// TwinCAT 3 PLC project PLC_Dyno
// ProgramVersion: 3.1.4026.25
// CompilerDefines: VISU_USEPROPERTYINFO
// libraries:
//   CmpBitmapPool, * (System)
//   Tc2_EtherCAT, * (Beckhoff Automation GmbH)
//   Tc2_MC2, * (Beckhoff Automation GmbH)
//   Tc2_MC2_Drive, * (Beckhoff Automation GmbH)
//   Tc2_Standard, * (Beckhoff Automation GmbH)
//   Tc2_System, * (Beckhoff Automation GmbH)
//   VisuDialogs, * (System)
//   VisuSymbols, 4.5.0.0 (System)
// project tree:
//   DUTs/ E_ControlMode.TcDUT, E_MotorState.TcDUT, E_SafetyState.TcTLEO, ST_AnalogInData.TcDUT, ST_EncoderData.TcDUT, ST_IOData.TcDUT, ST_MenteeMotorCmd.TcDUT, ST_MenteeMotorStatus.TcDUT, ST_MenteeMotorV32OsCmd.TcDUT, ST_MenteeMotorV32OsSample.TcDUT, ST_MenteeMotorV32OsStatus.TcDUT, ST_MenteeTrajCmd.TcDUT, ST_LoadProfileCmd.TcDUT, ST_CsvProfile.TcDUT, ST_Slot2Cfg.TcDUT, ST_MotorCommand.TcDUT, ST_RecChunk.TcDUT, U_WordReal.TcDUT, ST_MotorStatus.TcDUT, ST_Safety_Speps.TcDUT, ST_SyncSnapshot.TcDUT, ST_TwinSAFE_IN.TcDUT, ST_TwinSAFE_OUT.TcDUT, ST_UartBridgeCmd.TcDUT, ST_UartBridgeStatus.TcDUT
//   / GlobalTextList.TcGTLO, ImagePool.TcIPO (not stored), PlcTask.TcTTO, Visualization Manager.TcVMO (not stored), VISU_TASK.TcTTO
//   GVLs/ GVL_AnalogIn.TcGVL, GVL_Commands.TcGVL, GVL_MenteeFoe.TcGVL, GVL_Encoder.TcGVL, GVL_IO.TcGVL, GVL_MenteeMotor.TcGVL, GVL_MenteeMotorV32_OS.TcGVL, GVL_Profiles.TcGVL, GVL_CsvProfile.TcGVL, GVL_Slot2.TcGVL, GVL_Recording.TcGVL, GVL_Safety.TcGVL, GVL_Status.TcGVL, GVL_Sync.TcGVL, GVL_UartBridge.TcGVL
//   POUs/ CheckBounds.TcPOU, FB_AnalogInHandler.TcPOU, FB_EncoderHandler.TcPOU, FB_IOHandler.TcPOU, FB_MenteeMotorHandler.TcPOU, FB_MotorControl.TcPOU, FB_ExtSetpointProbe.TcPOU, FB_LoadMotorProfile.TcPOU, FB_CsvPlayer.TcPOU, FB_MenteeSdoCmd.TcPOU, FB_MenteeFoeFlash.TcPOU, FB_Slot2PipeHandler.TcPOU, FB_TorqueControl.TcPOU, FB_HighRateRecorder.TcPOU, FB_TrajectoryGen.TcPOU, FB_UartBridgeHandler.TcPOU, MAIN.TcPOU, PRG_Motion.TcPOU
//   VISUs/ Visualization.TcVIS
// real-time tasks:
//   TASK PlcTask: cycle T#1ms, priority 2, ADS port 350
//   TASK VISU_TASK: cycle T#200000us, priority 30, ADS port 351
// motion (NC):
//   TASK NC-Task 1 SAF: cycle T#1ms, priority 4, ADS port 501
//   TASK NC-Task 1 SVB: cycle T#10ms, priority 8, ADS port 511
//   AXIS Axis 1 (id 3)
//     General: UnitName=°
//     Dynamic: Acceleration=15000, Deceleration=15000, Jerk=178490.844
//     Velo: RefSearch=396.64632, RefSync=396.64632, SlowManual=1983.2316, FastManual=11899.3896, Fast=39664.632, Maximum=39664.632
//     OtherSettings: AllowMotionCmdToSlave=true
//     encoder EncType=8
//       EncPara: ScaleFactorNumerator=360, ScaleFactorDenominator=1048576, MaxCount=#xffffffff, EncPositionSource=1
//     drive DrvType=9
//       DrvPara: MaxCount=#xffffffff, DriveControlDWord=#x00030100
//         Analog: VeloReferenz=43631.0952, VeloScale=1.02400649589962, TorqueSetpointScale=10, ScaleFactorActTorque=0.1
//         TimeComp: TaskDelayCycles=1
//     controller CtrType=1
//       CtrPara: PriorControlFactor=1
//         Observer: BandWidth=20
//   AXIS Axis 2 (id 4)
//     General: UnitName=°
//     Dynamic: Acceleration=13437.441, Deceleration=13437.441, Jerk=40312.323
//     Velo: RefSearch=89.58294, RefSync=89.58294, SlowManual=447.9147, FastManual=2687.4882, Fast=8958.294, Maximum=8958.294
//     OtherSettings: AllowMotionCmdToSlave=true
//     encoder EncType=8
//       EncPara: ScaleFactorNumerator=360, ScaleFactorDenominator=1048576, MaxCount=#xffffffff
//     drive DrvType=9
//       DrvPara: MaxCount=#xffffffff, DriveControlDWord=#x00030100
//         Analog: VeloReferenz=9854.1234, VeloScale=1.02400649589962, TorqueSetpointScale=10, ScaleFactorActTorque=0.1
//         TimeComp: TaskDelayCycles=1
//     controller CtrType=1
//       CtrPara: PriorControlFactor=1
//         Observer: BandWidth=20
// I/O:
//   DEVICE Device 2 (EtherCAT), AmsNetId 192.168.1.50.3.1
//     Machine Side - A10 (EK1200)_1 [EK1200-5000 EtherCAT Power supply (2A E-Bus)]
//       A11 - DO (EL2022)_1 [EL2022 2Ch. Dig. Output 24V, 2A]
//       Term 3 (EL2502) [EL2502 2Ch. PWM output, 24V]
//       A12 - SI2 (EL1918)_1 [EL1918, 8Ch. Safety Input 24V, TwinSAFE]
//         modules: Module 1 (FSOE), Module 2 (FSLOGIC)
//       A13 - SO3 (EL2904)_1 [EL2904, 4 Ch. Safety Output 24V, 0.5A, TwinSAFE]
//         modules: Module 1 (FSOES), Module 2 (DO)
//       A14 - D-I/O (EL1859)_1 [EL1859 8Ch. Dig. Input 24V, 3ms, 8Ch. Dig. Output 24V, 0.5A]
//       A15 - AI (EL3002)_1 [EL3002 2Ch. Ana. Input +/-10V]
//       A19 - Enc (EL5112)_1 [EL5112 2Ch. Inc. Encoder 5V (2xAB or 1xABC RS422,TTL)]
//       A16 - AI  (EL3702)_1 [EL3702 2Ch. Ana. Input +/-10V, DIFF, Oversample]
//       A18 - Enc  (EL5112)_1 [EL5112 2Ch. Inc. Encoder 5V (2xAB or 1xABC RS422,TTL)]
//       A17 - AI  (EL3702)_1 [EL3702 2Ch. Ana. Input +/-10V, DIFF, Oversample]
//       Term 12 (EL5042) [EL5042 2Ch. BiSS-C Encoder]
//       Term 14 (EK1110)_1 [EK1110 EtherCAT extension]
//     Drive 1 (AX5112-0000-0216) [AX5112-0000-0216 EtherCAT Drive (SoE, 1 Ch.)]
//       STO_Drive1 (AX5805) [AX5805 (Safety Drive Option)]
//         modules: Module 1 (Safety Process Data, 1 axis), Module 2 (Standard Process Data, 1 axis)
//     Drive 2 (AX5125-0000-0216) [AX5125-0000-0216 EtherCAT Drive (SoE, 1 Ch.)]
//       STO_Drive2 (AX5805) [AX5805 (Safety Drive Option)]
//         modules: Module 1 (Safety Process Data, 1 axis), Module 2 (Standard Process Data, 1 axis)
//     Rack 19 (EK1100 - A0)_1 [EK1100 EtherCAT Coupler (2A E-Bus)]
//       A1 - SI1 (EL1918)_1 [EL1918, 8Ch. Safety Input 24V, TwinSAFE]
//         modules: Module 2 (FSLOGIC)
//       A2 -SO1 (EL2904)_1 [EL2904, 4 Ch. Safety Output 24V, 0.5A, TwinSAFE]
//         modules: Module 1 (FSOES), Module 2 (DO)
//       A3 - SO2 (EL2904)_1 [EL2904, 4 Ch. Safety Output 24V, 0.5A, TwinSAFE]
//         modules: Module 1 (FSOES), Module 2 (DO)
//       A4 - D-I/O (EL1859)_1 [EL1859 8Ch. Dig. Input 24V, 3ms, 8Ch. Dig. Output 24V, 0.5A]
//       A5 (EL9505)_1 [EL9505 Power supply terminal 5V]
//       A6  (EL9505)_1 [EL9505 Power supply terminal 5V]
//       Term 23 (EL9011) [EL9011 End Terminal]
//     Box 1 (Motor Slave) [Motor Slave]
// variable links:
//   Device 2 (EtherCAT) <-> Device 2 (EtherCAT)/Rack 19 (EK1100 - A0)_1/A1 - SI1 (EL1918)_1
//     Drive 1 (AX5112-0000-0216)/STO_Drive1 (AX5805)/Module 1 (Safety Process Data, 1 axis)/Inputs (Statusword)/FSOE <-> ConnectionOutputs/Message_71 RxPDO
//     Drive 2 (AX5125-0000-0216)/STO_Drive2 (AX5805)/Module 1 (Safety Process Data, 1 axis)/Inputs (Statusword)/FSOE <-> ConnectionOutputs/Message_72 RxPDO
//     Drive 1 (AX5112-0000-0216)/STO_Drive1 (AX5805)/Module 1 (Safety Process Data, 1 axis)/Outputs (Controlword)/FSOE <-> ConnectionInputs/Message_71 TxPDO
//     Drive 2 (AX5125-0000-0216)/STO_Drive2 (AX5805)/Module 1 (Safety Process Data, 1 axis)/Outputs (Controlword)/FSOE <-> ConnectionInputs/Message_72 TxPDO
//     Machine Side - A10 (EK1200)_1/A12 - SI2 (EL1918)_1/Module 1 (FSOE)/FSoE Inputs/FSOE <-> ConnectionOutputs/Message_62 RxPDO
//     Machine Side - A10 (EK1200)_1/A12 - SI2 (EL1918)_1/Module 1 (FSOE)/FSoE Outputs/FSOE <-> ConnectionInputs/Message_62 TxPDO
//     Machine Side - A10 (EK1200)_1/A13 - SO3 (EL2904)_1/Module 1 (FSOES)/RxPDO/FSOE <-> ConnectionInputs/Message_51 TxPDO
//     Machine Side - A10 (EK1200)_1/A13 - SO3 (EL2904)_1/Module 1 (FSOES)/TxPDO/FSOE <-> ConnectionOutputs/Message_51 RxPDO
//   Device 2 (EtherCAT) <-> Device 2 (EtherCAT)/Rack 19 (EK1100 - A0)_1/A2 -SO1 (EL2904)_1
//     Rack 19 (EK1100 - A0)_1/A1 - SI1 (EL1918)_1/ConnectionInputs/Message_7 TxPDO <-> Module 1 (FSOES)/RxPDO/FSOE
//     Rack 19 (EK1100 - A0)_1/A1 - SI1 (EL1918)_1/ConnectionOutputs/Message_7 RxPDO <-> Module 1 (FSOES)/TxPDO/FSOE
//   Device 2 (EtherCAT) <-> Device 2 (EtherCAT)/Rack 19 (EK1100 - A0)_1/A3 - SO2 (EL2904)_1
//     Rack 19 (EK1100 - A0)_1/A1 - SI1 (EL1918)_1/ConnectionInputs/Message_8 TxPDO <-> Module 1 (FSOES)/RxPDO/FSOE
//     Rack 19 (EK1100 - A0)_1/A1 - SI1 (EL1918)_1/ConnectionOutputs/Message_8 RxPDO <-> Module 1 (FSOES)/TxPDO/FSOE
//   NC-Task 1 SAF/Axes/Axis 1 <-> Device 2 (EtherCAT)/Drive 1 (AX5112-0000-0216)
//     Drive/Inputs/In/nDataIn1 <-> AT/Following distance
//     Drive/Inputs/In/nDataIn3[0] <-> AT/Torque/force feedback value
//     Drive/Inputs/In/nDcOutputTime <-> InfoData/DcOutputShift
//     Drive/Inputs/In/nState1 <-> AT/Drive status word @bit 8
//     Drive/Inputs/In/nState2 <-> AT/Drive status word
//     Drive/Inputs/In/nState4 @bit 1 <-> WcState/InputToggle
//     Drive/Inputs/In/nState4 <-> WcState/WcState
//     Drive/Outputs/Out/nCtrl1 <-> MDT/Master control word @bit 8
//     Drive/Outputs/Out/nDataOut1 <-> MDT/Position command value
//     Drive/Outputs/Out/nDataOut4[0] <-> MDT/Torque/force command value
//     Drive/Outputs/Out/nDataOut5 <-> MDT/High velocity limit value
//     Drive/Outputs/Out/nDataOut6 <-> MDT/Low velocity limit value
//     Enc/Inputs/In/nDataIn1 <-> AT/Position feedback 1 value
//     Enc/Inputs/In/nDataIn7 <-> AT/Velocity feedback 1 value
//     Enc/Inputs/In/nDcInputTime <-> InfoData/DcInputShift
//     Enc/Inputs/In/nState4 @bit 1 <-> WcState/InputToggle
//     Enc/Inputs/In/nState4 <-> WcState/WcState
//   NC-Task 1 SAF/Axes/Axis 2 <-> Device 2 (EtherCAT)/Drive 2 (AX5125-0000-0216)
//     Drive/Inputs/In/nDataIn1 <-> AT/Following distance
//     Drive/Inputs/In/nDcOutputTime <-> InfoData/DcOutputShift
//     Drive/Inputs/In/nState1 <-> AT/Drive status word @bit 8
//     Drive/Inputs/In/nState2 <-> AT/Drive status word
//     Drive/Inputs/In/nState4 @bit 1 <-> WcState/InputToggle
//     Drive/Inputs/In/nState4 <-> WcState/WcState
//     Drive/Outputs/Out/nCtrl1 <-> MDT/Master control word @bit 8
//     Drive/Outputs/Out/nDataOut1 <-> MDT/Position command value
//     Drive/Outputs/Out/nDataOut4[0] <-> MDT/Torque/force command value
//     Drive/Outputs/Out/nDataOut5 <-> MDT/High velocity limit value
//     Drive/Outputs/Out/nDataOut6 <-> MDT/Low velocity limit value
//     Enc/Inputs/In/nDataIn1 <-> AT/Position feedback 1 value
//     Enc/Inputs/In/nDcInputTime <-> InfoData/DcInputShift
//     Enc/Inputs/In/nState4 @bit 1 <-> WcState/InputToggle
//     Enc/Inputs/In/nState4 <-> WcState/WcState
//   PLC_Dyno/PLC_Dyno Instance <-> Device 2 (EtherCAT)/Box 1 (Motor Slave)
//     PlcTask Inputs/GVL_MenteeMotorV32_OS.nSlaveState <-> InfoData/State
//     PlcTask Inputs/PRG_Motion.fbMenteeSdo.stAdsAddr <-> InfoData/AdsAddr
//     PlcTask Inputs/PRG_Motion.fbSlot2Pipe.i_capture_count <-> Motor Response TB/capture_count
//     PlcTask Inputs/PRG_Motion.fbSlot2Pipe.i_categorial_error <-> Motor Response TB/categorial_error
//     PlcTask Inputs/PRG_Motion.fbSlot2Pipe.i_fault <-> Motor Response TB/fault
//     PlcTask Inputs/PRG_Motion.fbSlot2Pipe.i_fsm_state <-> Motor Response TB/fsm_state
//     PlcTask Inputs/PRG_Motion.fbSlot2Pipe.i_general_error <-> Motor Response TB/general_error
//     PlcTask Inputs/PRG_Motion.fbSlot2Pipe.i_last_op <-> Motor Response TB/last_op
//     PlcTask Inputs/PRG_Motion.fbSlot2Pipe.i_main_state <-> Motor Response TB/main_state
//     PlcTask Inputs/PRG_Motion.fbSlot2Pipe.i_motion_mode <-> Motor Response TB/motion_mode
//     PlcTask Inputs/PRG_Motion.fbSlot2Pipe.i_motor_enabled <-> Motor Response TB/motor_enabled
//     PlcTask Inputs/PRG_Motion.fbSlot2Pipe.i_sample_count <-> Motor Response TB/sample_count
//     PlcTask Inputs/PRG_Motion.fbSlot2Pipe.i_samples[{0..99}] <-> Motor Response TB/sample_{0..99}  (100 links)
//     PlcTask Inputs/PRG_Motion.fbSlot2Pipe.i_var_count <-> Motor Response TB/var_count
//     PlcTask Outputs/PRG_Motion.fbSlot2Pipe.q_addr <-> Motor Command TB/addr_payload
//     PlcTask Outputs/PRG_Motion.fbSlot2Pipe.q_inject[{0..9}] <-> Motor Command TB/inject_{0..9}  (10 links)
//     PlcTask Outputs/PRG_Motion.fbSlot2Pipe.q_op <-> Motor Command TB/op
//     PlcTask Outputs/PRG_Motion.fbSlot2Pipe.q_prescaler <-> Motor Command TB/prescaler
//     PlcTask Outputs/PRG_Motion.fbSlot2Pipe.q_size <-> Motor Command TB/size
//     PlcTask Outputs/PRG_Motion.fbSlot2Pipe.q_slot <-> Motor Command TB/slot
//     PlcTask Outputs/PRG_Motion.fbSlot2Pipe.q_strobe <-> Motor Command TB/strobe
//   PLC_Dyno/PLC_Dyno Instance <-> Device 2 (EtherCAT)/Drive 1 (AX5112-0000-0216)
//     PlcTask Inputs/PRG_Motion.fbMotor1.nActTorque_Raw <-> AT/Torque/force feedback value
//     PlcTask Outputs/GVL_Commands.nMotor1_CurrentLimit_Raw <-> MDT/Bipolar torque/force limit value
//   PLC_Dyno/PLC_Dyno Instance <-> Device 2 (EtherCAT)/Drive 2 (AX5125-0000-0216)
//     PlcTask Inputs/PRG_Motion.fbMotor2.nActTorque_Raw <-> AT/Torque/force feedback value
//     PlcTask Outputs/GVL_Commands.nMotor2_CurrentLimit_Raw <-> MDT/Bipolar torque/force limit value
//   PLC_Dyno/PLC_Dyno Instance <-> Device 2 (EtherCAT)/Machine Side - A10 (EK1200)_1/A14 - D-I/O (EL1859)_1
//     PlcTask Inputs/GVL_Safety.DoorMonitorFromPLC <-> Channel 2/Input
//     PlcTask Inputs/GVL_Safety.SolonoidStatus <-> Channel 1/Input
//     PlcTask Outputs/GVL_IO.BlueLED <-> Channel 11/Output
//     PlcTask Outputs/GVL_IO.GreenLED <-> Channel 10/Output
//     PlcTask Outputs/GVL_IO.RedLED <-> Channel 9/Output
//     PlcTask Outputs/GVL_IO.b_MotorCooling <-> Channel 12/Output
//   PLC_Dyno/PLC_Dyno Instance <-> Device 2 (EtherCAT)/Machine Side - A10 (EK1200)_1/A16 - AI  (EL3702)_1
//     PlcTask Inputs/PRG_Motion.fbAnalogIn1.nCh1_S{1..5} <-> Ch1 Sample {0..4}/Ch1 Value  (5 links)
//   PLC_Dyno/PLC_Dyno Instance <-> Device 2 (EtherCAT)/Machine Side - A10 (EK1200)_1/A17 - AI  (EL3702)_1
//     PlcTask Inputs/PRG_Motion.fbAnalogIn2.nCh1_S{1..5} <-> Ch1 Sample {0..4}/Ch1 Value  (5 links)
//   PLC_Dyno/PLC_Dyno Instance <-> Device 2 (EtherCAT)/Machine Side - A10 (EK1200)_1/A18 - Enc  (EL5112)_1
//     PlcTask Inputs/PRG_Motion.fbEncoder2.nCounterValue_Raw <-> ENC Status Channel 1/Counter value
//     PlcTask Inputs/PRG_Motion.fbEncoder2.nFrequencyValue_Raw <-> ENC Frequency Channel 1/Frequency value
//     PlcTask Outputs/PRG_Motion.fbEncoder2.nControlWord_Raw <-> ENC Control Channel 1/Control
//     PlcTask Outputs/PRG_Motion.fbEncoder2.nSetCounterValue_Raw <-> ENC Control Channel 1/Set counter value
//   PLC_Dyno/PLC_Dyno Instance <-> Device 2 (EtherCAT)/Machine Side - A10 (EK1200)_1/A19 - Enc (EL5112)_1
//     PlcTask Inputs/PRG_Motion.fbEncoder1.nCounterValue_Raw <-> ENC Status Channel 1/Counter value
//     PlcTask Inputs/PRG_Motion.fbEncoder1.nFrequencyValue_Raw <-> ENC Frequency Channel 1/Frequency value
//     PlcTask Outputs/PRG_Motion.fbEncoder1.nControlWord_Raw <-> ENC Control Channel 1/Control
//     PlcTask Outputs/PRG_Motion.fbEncoder1.nSetCounterValue_Raw <-> ENC Control Channel 1/Set counter value
//   PLC_Dyno/PLC_Dyno Instance <-> Device 2 (EtherCAT)/Rack 19 (EK1100 - A0)_1/A1 - SI1 (EL1918)_1
//     PlcTask Inputs/GVL_Safety.stTwinSAFE_IN/C1_FBK <-> StandardInputs/Standard Out Var 87
//     PlcTask Inputs/GVL_Safety.stTwinSAFE_IN/C2_FBK <-> StandardInputs/Standard Out Var 88
//     PlcTask Inputs/GVL_Safety.stTwinSAFE_IN/EStop_MantiRob <-> StandardInputs/Standard Out Var 84
//     PlcTask Inputs/GVL_Safety.stTwinSAFE_IN/EStop_NC1 <-> StandardInputs/Standard Out Var 82
//     PlcTask Inputs/GVL_Safety.stTwinSAFE_IN/EStop_NC2 <-> StandardInputs/Standard Out Var 83
//     PlcTask Inputs/GVL_Safety.stTwinSAFE_IN/EStop_Ok <-> StandardInputs/Standard Out Var 77
//     PlcTask Inputs/GVL_Safety.stTwinSAFE_IN/EStop_Status <-> StandardInputs/Standard Out Var 78
//     PlcTask Inputs/GVL_Safety.stTwinSAFE_IN/HV_Healthy <-> StandardInputs/Standard Out Var 90
//     PlcTask Inputs/GVL_Safety.stTwinSAFE_IN/HV_Interlock <-> StandardInputs/Standard Out Var 92
//     PlcTask Inputs/GVL_Safety.stTwinSAFE_IN/LV_Healthy <-> StandardInputs/Standard Out Var 89
//     PlcTask Inputs/GVL_Safety.stTwinSAFE_IN/LV_Interlock <-> StandardInputs/Standard Out Var 91
//     PlcTask Inputs/GVL_Safety.stTwinSAFE_IN/ReadyForStep2 <-> StandardInputs/Standard Out Var 52
//     PlcTask Inputs/GVL_Safety.stTwinSAFE_IN/STO_1 <-> StandardInputs/Standard Out Var 85
//     PlcTask Inputs/GVL_Safety.stTwinSAFE_IN/STO_2 <-> StandardInputs/Standard Out Var 86
//     PlcTask Inputs/GVL_Safety.stTwinSAFE_IN/Safety_Armed <-> StandardInputs/Standard Out Var 53
//     PlcTask Inputs/GVL_Safety.stTwinSAFE_IN/Speps/step{1..6} <-> StandardInputs/Standard Out Var {65..70}  (6 links)
//     PlcTask Inputs/GVL_Safety.stTwinSAFE_IN/Speps/stepRnD <-> StandardInputs/Standard Out Var 95
//     PlcTask Inputs/GVL_Safety.stTwinSAFE_IN/TransitionStep <-> StandardInputs/Standard Out Var 98
//     PlcTask Outputs/GVL_Safety.stTwinSAFE_OUT/BatRelay_Manual_Off <-> StandardOutputs/Standard In Var 56
//     PlcTask Outputs/GVL_Safety.stTwinSAFE_OUT/BatRelay_Manual_On <-> StandardOutputs/Standard In Var 55
//     PlcTask Outputs/GVL_Safety.stTwinSAFE_OUT/Bypass_C1C2 <-> StandardOutputs/Standard In Var 99
//     PlcTask Outputs/GVL_Safety.stTwinSAFE_OUT/DoorMonitor <-> StandardOutputs/Standard In Var 16
//     PlcTask Outputs/GVL_Safety.stTwinSAFE_OUT/ErrACK <-> StandardOutputs/Standard In Var 1
//     PlcTask Outputs/GVL_Safety.stTwinSAFE_OUT/EstopPLC <-> StandardOutputs/Standard In Var 54
//     PlcTask Outputs/GVL_Safety.stTwinSAFE_OUT/RB_BatBMS_Manual_Off <-> StandardOutputs/Standard In Var 58
//     PlcTask Outputs/GVL_Safety.stTwinSAFE_OUT/RB_BatBMS_Manual_On <-> StandardOutputs/Standard In Var 57
//     PlcTask Outputs/GVL_Safety.stTwinSAFE_OUT/RUN <-> StandardOutputs/Standard In Var 50
//     PlcTask Outputs/GVL_Safety.stTwinSAFE_OUT/Set_RnD_Mode <-> StandardOutputs/Standard In Var 94
//     PlcTask Outputs/GVL_Safety.stTwinSAFE_OUT/Set_RnD_Mode2 <-> StandardOutputs/Standard In Var 97
//     PlcTask Outputs/GVL_Safety.stTwinSAFE_OUT/SolenoedMonitor <-> StandardOutputs/Standard In Var 15
//   PLC_Dyno/PLC_Dyno Instance <-> NC-Task 1 SAF/Axes/Axis 1
//     PlcTask Inputs/PRG_Motion.Axis1.NcToPlc <-> Outputs/ToPlc
//     PlcTask Outputs/PRG_Motion.Axis1.PlcToNc <-> Inputs/FromPlc
//   PLC_Dyno/PLC_Dyno Instance <-> NC-Task 1 SAF/Axes/Axis 2
//     PlcTask Inputs/PRG_Motion.Axis2.NcToPlc <-> Outputs/ToPlc
//     PlcTask Outputs/PRG_Motion.Axis2.PlcToNc <-> Inputs/FromPlc

CONFIGURATION PLC_Dyno
    RESOURCE PLC ON TwinCAT3
        TASK PlcTask(INTERVAL := T#1ms, PRIORITY := 2);
        TASK VISU_TASK(INTERVAL := T#200000us, PRIORITY := 30);
        PROGRAM MAIN WITH PlcTask : MAIN;
        PROGRAM PRG_Motion WITH PlcTask : PRG_Motion;
        PROGRAM VisuElems_Visu_Prg WITH VISU_TASK : VisuElems.Visu_Prg;
    END_RESOURCE
END_CONFIGURATION

// ---- DUTs/E_ControlMode.TcDUT
TYPE E_ControlMode :
(
    IDLE        := 0,
    POSITION    := 1,
    VELOCITY    := 2,
    TORQUE      := 3
) UDINT := IDLE;
END_TYPE

// ---- DUTs/E_MotorState.TcDUT
TYPE E_MotorState :
(
    DISABLED    := 0,
    ENABLING    := 1,
    READY       := 2,
    MOVING      := 3,
    STOPPING    := 4,
    HOMING      := 5,
    ERROR       := 6,
    RESETTING   := 7    // sequenced fault recovery: SoE drive reset -> settle -> NC reset
) UDINT := DISABLED;
END_TYPE

// ---- DUTs/E_SafetyState.TcTLEO
{attribute 'qualified_only'}
{attribute 'strict'}
{attribute 'to_string'}
TYPE E_SafetyState :
(
	enum_RnD_2_Safe := 0,
	enum_Safe_2_RnD := 1,
	enum_RnD_2_Armed := 2,
	enum_Armed_2_RnD := 3
);
END_TYPE

// ---- DUTs/ST_AnalogInData.TcDUT
// EL3702 2-channel analog input with oversampling x5
// Written by FB_AnalogInHandler every cycle, read by Python via GVL_AnalogIn
TYPE ST_AnalogInData :
STRUCT
    //------------------------------------------------------------------
    // Raw oversampled inputs — 5 samples per channel per cycle
    // Linked to EL3702 PDOs in XAE (AT %I* in FB_AnalogInHandler)
    //------------------------------------------------------------------

    // Channel 1 — 5 oversamples [raw INT, -32768 to 32767]
    nCh1_Sample         : ARRAY[1..5] OF INT;

    // Channel 2 — 5 oversamples [raw INT, -32768 to 32767]
    nCh2_Sample         : ARRAY[1..5] OF INT;

    //------------------------------------------------------------------
    // Processed outputs — computed by FB_AnalogInHandler
    //------------------------------------------------------------------

    // Averaged value after oversampling processing [V]
    fCh1_Voltage        : LREAL;
    fCh2_Voltage        : LREAL;

    // Full scale range [V] — set once from MAIN (default ±10V)
    fFullScale          : LREAL := 10.0;

    // Status
    bError              : BOOL;
END_STRUCT
END_TYPE

// ---- DUTs/ST_EncoderData.TcDUT
TYPE ST_EncoderData :
STRUCT
    //------------------------------------------------------------------
    // Inputs — from EL5112 PDOs
    //------------------------------------------------------------------
    nStatusWord         : WORD;
    bInputA             : BOOL;
    bInputB             : BOOL;
    bInputC             : BOOL;
    bCounterUnderflow   : BOOL;
    bCounterOverflow    : BOOL;
    bLatchValid         : BOOL;
    bError              : BOOL;
    nCounterValue       : DWORD;
    nFrequencyValue     : DWORD;
    nState              : BYTE;
    fPosition           : LREAL;    // Scaled position [engineering units]

    //------------------------------------------------------------------
    // Outputs — written to EL5112 PDOs
    //------------------------------------------------------------------
    nSetCounterValue    : DWORD;    // Value to write to counter
    bSetCounter         : BOOL;     // Rising edge = write nSetCounterValue
    bZeroPosition       : BOOL;     // Rising edge = set counter to 0
END_STRUCT
END_TYPE

// ---- DUTs/ST_IOData.TcDUT
TYPE ST_IOData :
STRUCT
    //------------------------------------------------------------------
    // Digital inputs  (e.g. EL1008 — 8-channel 24V DC)
    //------------------------------------------------------------------

    // Raw 8-bit word from digital input terminal (bit 0 = DI channel 1)
    nDigitalInputs      : BYTE;

    // Named aliases — mapped in FB_IOHandler from nDigitalInputs bits
    bDI_EmergencyStop   : BOOL;   // Channel 1 — E-stop button
    bDI_HomeSensor_M1   : BOOL;   // Channel 2 — Home/ref switch Motor 1
    bDI_HomeSensor_M2   : BOOL;   // Channel 3 — Home/ref switch Motor 2
    bDI_LimitPos_M1     : BOOL;   // Channel 4 — Positive limit Motor 1
    bDI_LimitNeg_M1     : BOOL;   // Channel 5 — Negative limit Motor 1
    bDI_LimitPos_M2     : BOOL;   // Channel 6 — Positive limit Motor 2
    bDI_LimitNeg_M2     : BOOL;   // Channel 7 — Negative limit Motor 2
    bDI_UserInput1      : BOOL;   // Channel 8 — Spare / user-defined

    //------------------------------------------------------------------
    // Digital outputs  (e.g. EL2008 — 8-channel 24V DC)
    //------------------------------------------------------------------

    // Named aliases — written in FB_IOHandler, packed into nDigitalOutputs
    bDO_BrakeRelease_M1 : BOOL;   // Channel 1 — Release brake Motor 1
    bDO_BrakeRelease_M2 : BOOL;   // Channel 2 — Release brake Motor 2
    bDO_StatusLED_Green : BOOL;   // Channel 3 — System OK indicator
    bDO_StatusLED_Red   : BOOL;   // Channel 4 — Fault indicator
    bDO_UserOutput1     : BOOL;   // Channel 5 — Spare / user-defined
    bDO_UserOutput2     : BOOL;   // Channel 6 — Spare / user-defined

    // Packed output word (written to EL2008 terminal)
    nDigitalOutputs     : BYTE;

    //------------------------------------------------------------------
    // Analog inputs  (e.g. EL3002 — 2-channel ±10V or 0-20mA)
    //------------------------------------------------------------------

    // Raw ADC value from terminal [-32768 to 32767]
    nAnalogIn_Raw_Ch1   : INT;
    nAnalogIn_Raw_Ch2   : INT;

    // Scaled engineering values — conversion in FB_IOHandler
    fAnalogIn_Ch1       : LREAL;   // [V] or [mA] or user units
    fAnalogIn_Ch2       : LREAL;

    //------------------------------------------------------------------
    // Analog outputs  (e.g. EL4002 — 2-channel ±10V)
    //------------------------------------------------------------------

    // Setpoint from Python/GVL, written to terminal by FB_IOHandler
    fAnalogOut_Ch1      : LREAL;   // [V] or [mA] or user units
    fAnalogOut_Ch2      : LREAL;

    // Raw DAC value sent to terminal [-32768 to 32767]
    nAnalogOut_Raw_Ch1  : INT;
    nAnalogOut_Raw_Ch2  : INT;
END_STRUCT
END_TYPE

// ---- DUTs/ST_MenteeMotorCmd.TcDUT
// RxPDO — written by TwinCAT to Mentee Motor Slave (0x7000)
// Written by Python via GVL_MenteeMotor, consumed by FB_MenteeMotorHandler
TYPE ST_MenteeMotorCmd :
STRUCT
    kp                  : REAL;     // Position gain
    kd                  : REAL;     // Velocity gain
    p_des               : REAL;     // Desired position [rad or units]
    v_des               : REAL;     // Desired velocity [rad/s or units/s]
    torque_feed_forward : REAL;     // Feed forward torque [Nm or %]
    max_torque          : REAL;     // Max torque limit [Nm or %]
END_STRUCT
END_TYPE

// ---- DUTs/ST_MenteeMotorStatus.TcDUT
// TxPDO — read by TwinCAT from Mentee Motor Slave (0x6000)
// Written by FB_MenteeMotorHandler, read by Python via GVL_MenteeMotor
TYPE ST_MenteeMotorStatus :
STRUCT
    general_error_bits      : BYTE;     // General error flags
    categorial_error_bits   : BYTE;     // Categorical error flags
    motor_temp              : BYTE;     // Motor temperature [°C]
    theta                   : REAL;     // Actual position [rad or units]
    d_theta                 : REAL;     // Actual velocity [rad/s or units/s]
    measured_torque         : REAL;     // Measured torque [Nm or %]
    motor_torque_pi_in      : REAL;     // Torque PI controller input
    p_des_echo              : REAL;     // Echo of desired position setpoint
END_STRUCT
END_TYPE

// ---- DUTs/ST_MenteeMotorV32OsCmd.TcDUT
// RxPDO 0x1601 "Motor Command OS" — written by TwinCAT to Motor Slave V3.2 (0x7001)
// Written by Python via GVL_MenteeMotorV32_OS, consumed by FB_Slot2PipeHandler
TYPE ST_MenteeMotorV32OsCmd :
STRUCT
    nControlWord        : UDINT;    // 0x7001:01 control_word (raw 32-bit; packed per motor FW)
    impedance_p_des     : REAL;     // 0x7001:02 impedance_p_des
    impedance_v_des     : REAL;     // 0x7001:03 impedance_v_des
    impedance_kp        : REAL;     // 0x7001:04 impedance_kp
    impedance_kd        : REAL;     // 0x7001:05 impedance_kd
    impedance_torque_ff : REAL;     // 0x7001:06 impedance_torque_ff
    setpoint_position   : REAL;     // 0x7001:07 setpoint_position
    setpoint_velocity   : REAL;     // 0x7001:08 setpoint_velocity
    setpoint_current    : REAL;     // 0x7001:09 setpoint_current
    // Spare inject lanes 0/1/8/9 — RAW 32-bit values the app streams into the
    // matching q_inject slots (the FB copies them verbatim, NOT via the float
    // union). The app bit-encodes per the ELF-picked var's dtype (float bits vs
    // int). Slots 2..7 are the default command set (FW self-bound); these 4 are
    // free for ELF-picked inject targets.
    nRawInject0         : UDINT;    // -> q_inject[0]  (spare)
    nRawInject1         : UDINT;    // -> q_inject[1]  (spare)
    nRawInject8         : UDINT;    // -> q_inject[8]  (spare)
    nRawInject9         : UDINT;    // -> q_inject[9]  (spare)
END_STRUCT
END_TYPE

// ---- DUTs/ST_MenteeMotorV32OsSample.TcDUT
TYPE ST_MenteeMotorV32OsSample :
STRUCT
    // Generic oversample slot (flex-PDO 0x6001). w0/w1/w2 are RAW 32-bit words for
    // the fixed lanes:  w0=theta(F)  w1=d_theta(F)  w2=iq(F)
    sample_idx  : UDINT;    // sN_sample_idx — device oversample index
    w0          : UDINT;    // sN_w0 — raw word (float bits)
    w1          : UDINT;    // sN_w1
    w2          : UDINT;    // sN_w2
    // Extended lanes 3..9 — ELF-picked debug variables on the slot-2 debug
    // pipe. Filled by FB_Slot2PipeHandler from the SAME
    // capture index k as w0..w2 (the FW samples every bound lane on one
    // shared prescaler tick), so one aSamples[k] is one synchronized instant
    // stamped by sample_idx. Stay 0 when no debug var is bound to that lane.
    w3          : UDINT;
    w4          : UDINT;
    w5          : UDINT;
    w6          : UDINT;
    w7          : UDINT;
    w8          : UDINT;
    w9          : UDINT;
END_STRUCT
END_TYPE

// ---- DUTs/ST_MenteeMotorV32OsStatus.TcDUT
// TxPDO 0x1A01 "Motor Response OS" — read by TwinCAT from Motor Slave V3.2 (0x6001)
// Written by FB_Slot2PipeHandler, read by Python via GVL_MenteeMotorV32_OS / GVL_Sync snapshot
TYPE ST_MenteeMotorV32OsStatus :
STRUCT
    nStatusWord     : UDINT;                                    // 0x6001:01 status_word (raw)
    nSampleCount    : UDINT;                                    // 0x6001:02 sample_count (rolling)
    aSamples        : ARRAY[0..9] OF ST_MenteeMotorV32OsSample; // 0x6001:03..2A  s0..s9 buffer

    // Decoded status — V3.2 layout per MASTER_INTERFACE §4.4 (NOT the 3.1 bridge's)
    nFsmState               : BYTE;     // status_word bits 4:0  (fsm_state_e 0..19)
    nMainState              : BYTE;     // bits 8:5
    nOpMode                 : BYTE;     // bits 11:9 (MotionMode)
    nGroupId                : BYTE;     // DEPRECATED, always 0. The oversample-group
                                        // mechanism is gone (ELF debug-var lanes replaced
                                        // it) so nothing writes this. KEPT so the app's
                                        // by-name snapshot sum-read (which still lists the
                                        // field) can't break on activation order; drop it
                                        // together with that read.
    nGeneralErrorBits       : BYTE;     // bits 23:16
    nCategorialErrorBits    : BYTE;     // bits 31:24
    bError                  : BOOL;     // TRUE if any error bit set

    // Newest slot decoded as REAL (fixed lanes: w0/w1/w2 =
    // theta/d_theta/iq). Convenience for the trajectory anchor + the app's live
    // pos/vel/current readout (the app decodes the full slot stream per group).
    fLatestPos              : REAL;
    fLatestVel              : REAL;
    fLatestCurrent          : REAL;

    // EtherCAT AL state of the Motor Slave (from InfoData.State, set in
    // PRG_Motion). NOT from the TxPDO — it's the master's view of the slave.
    // Low nibble = AL state: 1=INIT, 2=PREOP, 4=SAFEOP, 8=OP; bit 4 (0x10) =
    // state error. The app treats (nAlState AND 16#000F) = 8 (OP) as connected.
    nAlState                : UINT;
END_STRUCT
END_TYPE

// ---- DUTs/ST_MenteeTrajCmd.TcDUT
// V3.2 generic motion-profile command + status, driven by FB_TrajectoryGen at
// the 1 kHz PLC task (profiling + injection are PLC-side; the app only configures
// + starts/stops). Profile shapes ported from the Cheetah mtb_serial_gui
// ProfileGenerator (Sinusoidal / Trapezoidal / Step / S-Curve / Ramp), evaluated
// online as value(t). The selected field (nField) is driven while running.
// Position/Impedance profiles are anchored at the rotor's current position
// (added as an offset) so they never jump at Start; Velocity/Current are absolute.
// ADS symbol: GVL_MenteeMotorV32_OS.stTraj
TYPE ST_MenteeTrajCmd :
STRUCT
    // --- selection ---
    nShape       : BYTE;    // 0 Sinusoidal | 1 Trapezoidal | 2 Step | 3 S-Curve | 4 Ramp
    nField       : BYTE;    // 0 setpoint_position | 1 impedance_p_des | 2 setpoint_velocity | 3 setpoint_current

    // --- shape parameters (union; only the relevant ones are used per shape) ---
    fAmplitude   : REAL;    // Sinusoidal
    fFrequency   : REAL;    // Sinusoidal [Hz]
    fOffset      : REAL;    // Sinusoidal
    fStartValue  : REAL;    // Trapezoid/S-Curve/Ramp start; Step initial
    fPeakValue   : REAL;    // Trapezoid/S-Curve peak
    fEndValue    : REAL;    // Ramp end; Step final
    fAccelTime   : REAL;    // Trapezoid/S-Curve ramp-up [s]
    fSteadyTime  : REAL;    // Trapezoid/S-Curve hold [s]
    fDecelTime   : REAL;    // Trapezoid/S-Curve ramp-down [s]
    fStepTime    : REAL;    // Step transition time [s]
    fDuration    : REAL;    // Sinusoidal/Step/Ramp total time [s]

    // --- repeat (loop the whole profile) ---
    bRepetitive  : BOOL;
    nReps        : UDINT;   // 0 = infinite
    fRestS       : REAL;    // rest between reps [s]

    // --- control ---
    bStart       : BOOL;    // rising edge -> (re)start
    bStop        : BOOL;    // rising edge -> abort + hold

    // --- status (written by FB_TrajectoryGen) ---
    bRunning     : BOOL;
    fSetpoint    : REAL;    // current generated setpoint
    fElapsed     : REAL;    // elapsed time in the current run [s]
END_STRUCT
END_TYPE

// ---- DUTs/ST_LoadProfileCmd.TcDUT
// Load-motor (Beckhoff AX5000) motion-profile command + status, driven by
// FB_LoadMotorProfile at the PLC task rate. Same online value(t) shapes as
// ST_MenteeTrajCmd / FB_TrajectoryGen (Sinusoidal / Trapezoidal / Step /
// S-Curve / Ramp), but with a DOMAIN selector because a load motor can run the
// profile as a TORQUE waveform (streamed into the existing MC_TorqueControl via
// stMotorN_Cmd.fTargetTorque) or as a POSITION / VELOCITY waveform (external
// setpoint generation MC_ExtSetPointGen* on the NC axis).
//
// Values are in PLC-native units (the backend pre-converts): TORQUE = % of motor
// rated; POSITION = deg; VELOCITY = deg/s (gear-scaled). Position profiles anchor
// at the axis actual position at Start (no jump); velocity integrates to position
// for the external-setpoint feed; torque is absolute.
//
// One per load motor in GVL_Profiles (stLoadProfile1 / stLoadProfile2). Started
// either directly (bStart) or, for a synchronized run, by GVL_Profiles.bStartSync
// (gated by bEnable) so it begins on the exact same PLC cycle as the Mentee half.
TYPE ST_LoadProfileCmd :
STRUCT
    // --- domain + selection ---
    nDomain      : BYTE;    // 0 TORQUE (-> fTargetTorque) | 1 POSITION | 2 VELOCITY (ext-setpoint)
    nShape       : BYTE;    // 0 Sinusoidal | 1 Trapezoidal | 2 Step | 3 S-Curve | 4 Ramp

    // --- shape parameters (union; only the relevant ones are used per shape) ---
    fAmplitude   : REAL;    // Sinusoidal
    fFrequency   : REAL;    // Sinusoidal [Hz]
    fOffset      : REAL;    // Sinusoidal
    fStartValue  : REAL;    // Trapezoid/S-Curve/Ramp start; Step initial
    fPeakValue   : REAL;    // Trapezoid/S-Curve peak
    fEndValue    : REAL;    // Ramp end; Step final
    fAccelTime   : REAL;    // Trapezoid/S-Curve ramp-up [s]
    fSteadyTime  : REAL;    // Trapezoid/S-Curve hold [s]
    fDecelTime   : REAL;    // Trapezoid/S-Curve ramp-down [s]
    fStepTime    : REAL;    // Step transition time [s]
    fDuration    : REAL;    // Sinusoidal/Step/Ramp total time [s]

    // --- repeat (loop the whole profile) ---
    bRepetitive  : BOOL;
    nReps        : UDINT;   // 0 = infinite
    fRestS       : REAL;    // rest between reps [s]

    // --- control ---
    bEnable      : BOOL;    // participate in a synchronized (bStartSync) run
    bStart       : BOOL;    // rising edge -> (re)start this profile alone
    bStop        : BOOL;    // rising edge -> abort + hold

    // --- status (written by FB_LoadMotorProfile) ---
    bRunning     : BOOL;
    bExtActive   : BOOL;    // POSITION/VELOCITY: external setpoint generator engaged
    fSetpoint    : REAL;    // current generated value (native units)
    fElapsed     : REAL;    // elapsed time in the current run [s]
END_STRUCT
END_TYPE

// ---- DUTs/ST_CsvProfile.TcDUT
// Generic CSV-trajectory buffer + config, replayed by FB_CsvPlayer at the task
// rate. The app parses a CSV (time, mentee setpoint, beckhoff setpoint), resamples
// it to a uniform period, converts each USED channel to PLC-native units, uploads
// the sample arrays here, sets nCount/fSampleDt + the per-motor selectors, then
// pulses bStart. FB_CsvPlayer steps through the buffer by elapsed time (linear
// interpolation), emitting BOTH setpoints from the same time index -> the two
// motors are inherently synchronized (one player, one clock).
//
// Values are ABSOLUTE (no anchoring): mentee position/velocity/current and beckhoff
// torque/position/velocity are commanded as the literal (converted) sample values.
// => a position run jumps to sample 0 at start if the motor isn't already there.
//
// The array bound below is the SINGLE SOURCE OF TRUTH for the buffer capacity: the
// app reads this array's byte size live over ADS (backend motor_service._csv_capacity)
// and adapts its row cap + duration preview automatically, so resizing here needs NO
// app-code change. 300000 samples = 300 s @ 1 kHz (or longer at a coarser fSampleDt;
// the player interpolates back up to the task rate). aMentee/aLoad are REAL (native
// units after conversion); at 300000 the two buffers are ~2.4 MB (fits the data area).
TYPE ST_CsvProfile :
STRUCT
    // --- sample buffers (filled by the app BEFORE bStart) ---
    aMentee       : ARRAY[0..299999] OF REAL;  // mentee setpoint samples (native units)
    aLoad         : ARRAY[0..299999] OF REAL;  // beckhoff setpoint samples (native units)
    nCount        : UDINT;     // number of valid samples in each array (<= array bound)
    fSampleDt     : REAL;      // uniform sample period [s]

    // --- mentee selection ---
    bMenteeEnable : BOOL;      // drive the Mentee from aMentee
    nMenteeField  : BYTE;      // 0 setpoint_position | 1 impedance_p_des | 2 setpoint_velocity | 3 setpoint_current

    // --- beckhoff selection ---
    bLoadEnable   : BOOL;      // drive a load motor from aLoad
    nLoadMotor    : BYTE;      // 1 or 2 (which load axis)
    nLoadDomain   : BYTE;      // 0 TORQUE (-> fTargetTorque) | 1 POSITION | 2 VELOCITY (ext-setpoint)

    // --- repeat (loop the whole table) ---
    bRepetitive   : BOOL;
    nReps         : UDINT;     // 0 = infinite
    fRestS        : REAL;      // rest between reps [s]

    // --- control ---
    bStart        : BOOL;      // rising edge -> (re)play from sample 0 (latches the scalar config)
    bStop         : BOOL;      // rising edge -> abort + hold

    // --- status (written by FB_CsvPlayer) ---
    bRunning      : BOOL;
    bLoadExtActive: BOOL;      // POSITION/VELOCITY: external setpoint generator engaged
    fElapsed      : REAL;      // elapsed time in the current pass [s]
    fMenteeOut    : REAL;      // current interpolated mentee value (native units)
    fLoadOut      : REAL;      // current interpolated load value (native units)
END_STRUCT
END_TYPE

// ---- DUTs/ST_Slot2Cfg.TcDUT
// Binding configuration for the generic slot-2 debug PDO pipe (SLOT2_DEBUG_PDO_PROTOCOL).
// The app fills the ABSOLUTE slave RAM addresses (from the flashed FW build's .map/.elf —
// they move every build!) and pulses GVL_Slot2.bConfigure; FB_Slot2PipeHandler then walks
// the table over the op/strobe protocol (CLEAR_ALL, then one bind per entry with addr<>0).
//
// Fixed conventions (mirror the app config + the old fixed pipe):
//   monitor lanes: 0=theta  1=d_theta  2=iq  |  3..9 = ELF-picked debug variables
//   inject slots: 0=impedance_p_des 1=impedance_v_des 2=impedance_kp 3=impedance_kd
//                 4=impedance_torque_ff 5=setpoint_position 6=setpoint_velocity 7=setpoint_current
TYPE ST_Slot2Cfg :
STRUCT
    aMonAddr    : ARRAY[0..9] OF UDINT;   // monitor lane -> absolute RAM addr (0 = unbound)
    aMonSize    : ARRAY[0..9] OF UDINT;   // width code: 0=1B, 1=2B, else 4B (default 4B)
    aInjAddr    : ARRAY[0..9] OF UDINT;   // inject slot -> absolute RAM addr (0 = unbound)
    aInjSize    : ARRAY[0..9] OF UDINT;
    nPrescaler  : UDINT := 5;             // capture decimation (40 kHz / prescaler; 5 -> 8 kHz,
                                          // 8 samples per 1 ms cycle = 20% headroom, no drops)
    nProfileId  : BYTE;                   // DEPRECATED, unused. Was the oversample-group
                                          // selector; that mechanism is gone. KEPT because
                                          // the app still writes 0 here (pinning the group
                                          // off on older PLC builds) — deleting it before
                                          // that write would fail every bind. Drop both
                                          // together.
END_STRUCT
END_TYPE

// ---- DUTs/ST_MotorCommand.TcDUT
TYPE ST_MotorCommand :
STRUCT
    //------------------------------------------------------------------
    // Control
    //------------------------------------------------------------------
    bEnable             : BOOL;         // TRUE = enable drive power
    bResetError         : BOOL;         // Rising edge = reset active fault (sequenced:
                                        // SoE drive reset -> 250 ms settle -> NC reset)
    bSoeReset           : BOOL;         // Rising edge = SoE drive reset ONLY (S-0-0099,
                                        // diagnostic; runs in background from any state)
    bNcReset            : BOOL;         // Rising edge = NC axis reset ONLY (MC_Reset,
                                        // diagnostic; runs in background from any state)
    bHome               : BOOL;         // Rising edge = start homing sequence
    bStop               : BOOL;         // Rising edge = decelerate to standstill
    bZeroPosition       : BOOL;         // Rising edge = set current position to 0
    eControlMode        : E_ControlMode;

    //------------------------------------------------------------------
    // Position mode  (eControlMode = POSITION)
    //------------------------------------------------------------------
    fTargetPosition     : LREAL;        // Target position [units]
    fDirection          : LREAL := 1.0; // Move direction for relative moves
    bRelative           : BOOL;         // TRUE = relative, FALSE = absolute
    bExecuteMove        : BOOL;         // Rising edge = execute move

    //------------------------------------------------------------------
    // Velocity mode  (eControlMode = VELOCITY)
    //------------------------------------------------------------------
    fTargetVelocity     : LREAL;        // Target velocity [units/s] sign = direction

    //------------------------------------------------------------------
    // Torque mode  (FB_TorqueControl)
    //------------------------------------------------------------------
    bTorqueExecute      : BOOL;         // Hold TRUE = torque active, FALSE = stop
    fTargetTorque       : LREAL;        // Target torque [% of rated, -100 to 100]
    fTorqueRamp         : LREAL := 100.0; // Torque ramp [% / s]
    fTorqueVelLimitHigh : LREAL := 859.437;  // Velocity safety limit [deg/s] = 15 rad/s
    fTorqueVelLimitLow  : LREAL := -859.437; // = -15 rad/s

    //------------------------------------------------------------------
    // Motion profile (shared across position and velocity modes)
    //------------------------------------------------------------------
    fAcceleration       : LREAL := 500.0;
    fDeceleration       : LREAL := 500.0;
    fJerk               : LREAL := 0.0;
    fMaxVelocity        : LREAL := 100.0;

    //------------------------------------------------------------------
    // Drive current/torque limit -> AX5000 SoE S-0-0092 (applies in all modes,
    // incl. position mode S-0-0032 = 11). Scaled to the PDO in PRG_Motion.
    //------------------------------------------------------------------
    fCurrentLimit_pct   : LREAL := 100.0; // [%] 0..100 of motor peak (P-0-0092)
END_STRUCT
END_TYPE

// ---- DUTs/ST_RecChunk.TcDUT
// High-rate recording chunk — struct-of-arrays (SoA) so the app can bulk-read
// each channel as a flat typed array over ADS (no struct packing/alignment).
//
// One CHUNK = REC_CHUNK EtherCAT frames. The recorder FB fills the active chunk
// one frame per cycle; when full it advances to the next chunk in the ring and
// bumps GVL_Recording.nChunkSeq. The app reads each completed chunk's arrays in
// one bulk ADS read per channel, then writes them to the recording file.
//
// Two rates share one DC timebase:
//   * bus-rate  (one value per frame): aDcTs + load motors / Futek / Mentee status
//   * Mentee    (REC_OVERSAMPLE per frame): aMn* arrays, length REC_CHUNK*REC_OVERSAMPLE
//
// Sizes are compile-time constants in GVL_Recording — keep them in lock-step
// with the FB and the backend reader (chunk length + oversample count).
TYPE ST_RecChunk :
STRUCT
    nCount   : UDINT;   // frames actually filled in this chunk (= REC_CHUNK when complete)

    // ── bus-rate channels (one element per frame) ──────────────────────
    // Types match the source snapshot fields exactly (no implicit conversion):
    // load motors / analog are LREAL; encoder counters are DWORD.
    aDcTs    : ARRAY[0..GVL_Recording.REC_CHUNK - 1] OF ULINT;   // DC time, 100 ns ticks
    aM1Pos   : ARRAY[0..GVL_Recording.REC_CHUNK - 1] OF LREAL;   // load motor 1
    aM1Vel   : ARRAY[0..GVL_Recording.REC_CHUNK - 1] OF LREAL;
    aM1Trq   : ARRAY[0..GVL_Recording.REC_CHUNK - 1] OF LREAL;
    aM2Pos   : ARRAY[0..GVL_Recording.REC_CHUNK - 1] OF LREAL;   // load motor 2
    aM2Vel   : ARRAY[0..GVL_Recording.REC_CHUNK - 1] OF LREAL;
    aM2Trq   : ARRAY[0..GVL_Recording.REC_CHUNK - 1] OF LREAL;
    aEnc1Cnt : ARRAY[0..GVL_Recording.REC_CHUNK - 1] OF DWORD;   // Futek 1 encoder
    aEnc1Frq : ARRAY[0..GVL_Recording.REC_CHUNK - 1] OF DWORD;
    aEnc2Cnt : ARRAY[0..GVL_Recording.REC_CHUNK - 1] OF DWORD;   // Futek 2 encoder
    aEnc2Frq : ARRAY[0..GVL_Recording.REC_CHUNK - 1] OF DWORD;
    aAin1V   : ARRAY[0..GVL_Recording.REC_CHUNK - 1] OF LREAL;   // Futek 1 analog (V)
    aAin2V   : ARRAY[0..GVL_Recording.REC_CHUNK - 1] OF LREAL;   // Futek 2 analog (V)
    aMnSW    : ARRAY[0..GVL_Recording.REC_CHUNK - 1] OF UDINT;   // Mentee status word (bus-rate)
    aMnCnt   : ARRAY[0..GVL_Recording.REC_CHUNK - 1] OF UDINT;   // fresh oversamples this frame (0..REC_OVERSAMPLE)

    // ── Mentee oversamples (REC_OVERSAMPLE per frame) — raw slot words ──
    // w0/w1/w2 are raw 32-bit words for the fixed lanes (theta / d_theta / iq).
    // Storing them raw keeps the recorder decode-agnostic — the app reinterprets
    // the bits per lane.
    aMnIdx   : ARRAY[0..GVL_Recording.REC_CHUNK * GVL_Recording.REC_OVERSAMPLE - 1] OF UDINT; // sample_idx
    aMnW0    : ARRAY[0..GVL_Recording.REC_CHUNK * GVL_Recording.REC_OVERSAMPLE - 1] OF UDINT;
    aMnW1    : ARRAY[0..GVL_Recording.REC_CHUNK * GVL_Recording.REC_OVERSAMPLE - 1] OF UDINT;
    aMnW2    : ARRAY[0..GVL_Recording.REC_CHUNK * GVL_Recording.REC_OVERSAMPLE - 1] OF UDINT;
    // ── extended lanes 3..9 — ELF-picked debug variables (slot-2 pipe) ──
    // Same flat index as aMnIdx/aMnW0..2 (frame*REC_OVERSAMPLE + slot), so
    // element i of EVERY aMn* array is the same synchronized capture instant.
    // Kept LAST so the app can skip reading them when nothing is selected.
    aMnW3    : ARRAY[0..GVL_Recording.REC_CHUNK * GVL_Recording.REC_OVERSAMPLE - 1] OF UDINT;
    aMnW4    : ARRAY[0..GVL_Recording.REC_CHUNK * GVL_Recording.REC_OVERSAMPLE - 1] OF UDINT;
    aMnW5    : ARRAY[0..GVL_Recording.REC_CHUNK * GVL_Recording.REC_OVERSAMPLE - 1] OF UDINT;
    aMnW6    : ARRAY[0..GVL_Recording.REC_CHUNK * GVL_Recording.REC_OVERSAMPLE - 1] OF UDINT;
    aMnW7    : ARRAY[0..GVL_Recording.REC_CHUNK * GVL_Recording.REC_OVERSAMPLE - 1] OF UDINT;
    aMnW8    : ARRAY[0..GVL_Recording.REC_CHUNK * GVL_Recording.REC_OVERSAMPLE - 1] OF UDINT;
    aMnW9    : ARRAY[0..GVL_Recording.REC_CHUNK * GVL_Recording.REC_OVERSAMPLE - 1] OF UDINT;

    // ── Futek analog oversamples (REC_FUTEK_OS per frame) — EL3702 x5, in Volts ──
    // Flat index frame*REC_FUTEK_OS + slot. Stored as V (same scale as aAin1V) so
    // the backend's volts->Nm calibration path handles them identically, at 5x rate.
    aFut1V   : ARRAY[0..GVL_Recording.REC_CHUNK * GVL_Recording.REC_FUTEK_OS - 1] OF LREAL;   // Futek 1 (stAnalogIn1 ch1)
    aFut2V   : ARRAY[0..GVL_Recording.REC_CHUNK * GVL_Recording.REC_FUTEK_OS - 1] OF LREAL;   // Futek 2 (stAnalogIn2 ch1)
END_STRUCT
END_TYPE

// ---- DUTs/U_WordReal.TcDUT
// Bit-reinterpret a raw 32-bit oversample word (UDINT on the wire) as IEEE-754
// REAL — the flex-PDO slot words are float-bits for the motion/iq fields.
TYPE U_WordReal :
UNION
    u : UDINT;
    f : REAL;
END_UNION
END_TYPE

// ---- DUTs/ST_MotorStatus.TcDUT
TYPE ST_MotorStatus :
STRUCT
    //------------------------------------------------------------------
    // State machine
    //------------------------------------------------------------------
    eState              : E_MotorState;
    eControlMode        : E_ControlMode;

    //------------------------------------------------------------------
    // Status flags
    //------------------------------------------------------------------
    bEnabled            : BOOL;     // Drive power is on and ready
    bMoving             : BOOL;     // Axis is in motion
    bAtTarget           : BOOL;     // Position/velocity within tolerance
    bHomingDone         : BOOL;     // Homing completed successfully
    bZeroDone           : BOOL;     // Zero position completed successfully
    bTorqueActive       : BOOL;     // Torque control is active
    bTorqueInTorque     : BOOL;     // Target torque reached
    bError              : BOOL;     // Fault active
    nErrorID            : UDINT;    // TwinCAT NC error code (0 = no error)
    nResetStage         : BYTE;     // fault-recovery progress: 0 idle | 1 SoE drive
                                    // reset | 2 settle | 3 NC reset

    //------------------------------------------------------------------
    // Actual values
    //------------------------------------------------------------------
    fActPosition        : LREAL;    // [units]
    fActVelocity        : LREAL;    // [units/s]
    fActTorque          : LREAL;    // [% of rated torque]

    //------------------------------------------------------------------
    // Diagnostics
    //------------------------------------------------------------------
    fDcBusVoltage       : LREAL;    // [V]  — requires drive PDO mapping
    fDriveTemp          : LREAL;    // [°C] — requires drive PDO mapping
    nTimestamp          : UDINT;    // [ms since PLC start]
END_STRUCT
END_TYPE

// ---- DUTs/ST_Safety_Speps.TcDUT
TYPE ST_Safety_Speps :
STRUCT
	step1: BOOL;
	step2: BOOL;
	step3: BOOL;
	step4: BOOL;
	step5: BOOL;
	step6: BOOL;
	stepRnD	:	BOOL	;

END_STRUCT
END_TYPE

// ---- DUTs/ST_SyncSnapshot.TcDUT
TYPE ST_SyncSnapshot :
STRUCT
    // Cycle identification
    nCycleCount             : UDINT;    // Increments each PLC cycle
    nDcTimestamp            : ULINT;    // DC time in nanoseconds (F_GetCurDcTaskTime64 / DCTIME64)

    // UART Bridge — V3.1 status + live data
    stBridge                : ST_UartBridgeStatus;

    // Mentee Motor — V3.2 direct motor status
    stMotor                 : ST_MenteeMotorStatus;

    // Encoders
    stEncoder1              : ST_EncoderData;
    stEncoder2              : ST_EncoderData;

    // Analog inputs
    stAnalogIn1             : ST_AnalogInData;
    stAnalogIn2             : ST_AnalogInData;

    // Motor control status
    stMotor1Status          : ST_MotorStatus;
    stMotor2Status          : ST_MotorStatus;

    // Safety
    bEStopActive            : BOOL;
	
	stMotorV32_OS           : ST_MenteeMotorV32OsStatus;    // V3.2 motor #2 (slot-2 OS, 0x1A01)  <-- NEW
	bTrajRunning            : BOOL;                         // V3.2 trajectory generator active (FB_TrajectoryGen)
END_STRUCT
END_TYPE

// ---- DUTs/ST_TwinSAFE_IN.TcDUT
TYPE ST_TwinSAFE_IN :
STRUCT
	Safety_Armed: BOOL;
	ReadyForStep2: BOOL;
	Speps: ST_Safety_Speps;
	EStop_Ok	:	BOOL	;//SI 2026 05 25
	EStop_Status:	BOOL	;//SI 2026 05 25
	TransitionStep	:	BOOL	;
	

	EStop_NC1	:	BOOL	;
	EStop_NC2	:	BOOL	;
	EStop_MantiRob : BOOL	;
	STO_1		:	BOOL	;
	STO_2		:	BOOL	;
	C1_FBK		:	BOOL	;
	C2_FBK		:	BOOL	;
	LV_Healthy	:	BOOL	;
	HV_Healthy	:	BOOL	;
	
	LV_Healthy_Invert	:	BOOL	;
	HV_Healthy_Invert	:	BOOL	;
	
	LV_Interlock	:	BOOL	;
	HV_Interlock	:	BOOL	;

END_STRUCT
END_TYPE

// ---- DUTs/ST_TwinSAFE_OUT.TcDUT
TYPE ST_TwinSAFE_OUT :
STRUCT
	
	RUN			: BOOL := TRUE;
	ErrACK		: BOOL:=TRUE;
	Restart		: BOOL;
	DoorMonitor: BOOL;
	SolenoedMonitor: BOOL;

	BatRelay_CMD: BOOL;
	BatRelay_Manual_Off: BOOL;
	BatRelay_Manual_On: BOOL;
	Set_RnD_Mode	:	BOOL	;
	Set_RnD_Mode2	:	BOOL	;

	EstopPLC: BOOL;

	BatBMS_Cmd: BOOL;
	RB_BatBMS_Manual_Off: BOOL;
	RB_BatBMS_Manual_On: BOOL;
	Bypass_C1C2	:	BOOL	;

END_STRUCT
END_TYPE

// ---- DUTs/ST_UartBridgeCmd.TcDUT
// RxPDO — written by TwinCAT to UART Bridge Slave (0x7000)
TYPE ST_UartBridgeCmd :
STRUCT
    //------------------------------------------------------------------
    // Control word — packed by FB_UartBridgeHandler from named bits below
    // Bit 0:     arm           (rising edge)
    // Bit 1:     idle          (rising edge)
    // Bit 2:     gate_block    (rising edge)
    // Bit 3:     calibrate     (rising edge)
    // Bit 4:     bode          (rising edge)
    // Bit 5:     noodle        (rising edge)
    // Bit 6:     reset         (rising edge)
    // Bit 7:     led_on        (rising edge)
    // Bit 8:     led_off       (rising edge)
    // Bit 9:     query_state   (rising edge)
    // Bits 11:10 bridge_mode   (level: 0=OFF, 1=MONITOR, 2=RECORDING)
    // Bits 14:12 motion_mode   (level: 0=Noodle, 1=Pos, 2=Vel, 3=Torque, 4=Impedance)
    //------------------------------------------------------------------

    // Rising edge commands — pulse TRUE then FALSE from Python
    bArm            : BOOL;
    bIdle           : BOOL;
    bGateBlock      : BOOL;
    bCalibrate      : BOOL;
    bBode           : BOOL;
    bNoodle         : BOOL;
    bReset          : BOOL;
    bLedOn          : BOOL;
    bLedOff         : BOOL;
    bQueryState     : BOOL;

    // Level commands
    nBridgeMode     : BYTE := 1;    // 0=OFF, 1=MONITOR, 2=RECORDING — default MONITOR
    nMotionMode     : BYTE;     // 0=Noodle, 1=Pos, 2=Vel, 3=Torque, 4=Impedance

    // Motion parameters
    p_des           : REAL;     // Desired position
    v_des           : REAL;     // Desired velocity
    kp              : REAL;     // Position gain
    kd              : REAL;     // Velocity gain
    torque_ff       : REAL;     // Feed forward torque
END_STRUCT
END_TYPE

// ---- DUTs/ST_UartBridgeStatus.TcDUT
// TxPDO — read by TwinCAT from UART Bridge Slave (0x6000)
TYPE ST_UartBridgeStatus :
STRUCT
    //------------------------------------------------------------------
    // Status word — decoded by FB_UartBridgeHandler
    // Bits 3:0:   fsm_state
    // Bits 7:4:   main_state
    // Bits 10:8:  op_mode
    // Bits 12:11: bridge_mode (echo)
    // Bits 23:16: general_error_bits
    // Bits 31:24: categorial_error_bits
    //------------------------------------------------------------------
    nStatusWord             : UDINT;    // Raw status word

    // Decoded status fields
    nFsmState               : BYTE;     // Bits 3:0
    nMainState              : BYTE;     // Bits 7:4
    nOpMode                 : BYTE;     // Bits 10:8
    nBridgeModeEcho         : BYTE;     // Bits 12:11
    nGeneralErrorBits       : BYTE;     // Bits 23:16
    nCategorialErrorBits    : BYTE;     // Bits 31:24
    bError                  : BOOL;     // TRUE if any error bit set

    // Diagnostics
    nPacketCount            : UINT;     // Rolling packet counter
    nTimestamp              : UDINT;    // Device timestamp

    // Live V3.1 data
    bldc_pos                : REAL;     // BLDC actual position
    filtered_p_des          : REAL;     // Filtered position setpoint
    bldc_vel                : REAL;     // BLDC actual velocity
    v_des                   : REAL;     // Velocity setpoint echo
    measured_current        : REAL;     // Measured motor current
    p_i_input               : REAL;     // PI controller input
    impedance_output        : REAL;     // Impedance controller output
END_STRUCT
END_TYPE

// ---- GVLs/GVL_AnalogIn.TcGVL
{attribute 'TcGvlVarFlags' := 'OPC'}
VAR_GLOBAL
    // EL3702 analog input data — written by FB_AnalogInHandler, read by Python over ADS
    // ADS symbol: GVL_AnalogIn.stAnalogIn
    stAnalogIn1         : ST_AnalogInData;
    stAnalogIn2         : ST_AnalogInData;
END_VAR

// ---- GVLs/GVL_Commands.TcGVL
VAR_GLOBAL
    // GVL_Commands — motor command interface written by Python over ADS, plus the
    // AX5000 current/torque-limit PDO outputs. ADS symbols: GVL_Commands.stMotor1_Cmd
    //                                                        GVL_Commands.stMotor2_Cmd
    stMotor1_Cmd    : ST_MotorCommand;
    stMotor2_Cmd    : ST_MotorCommand;

    // AX5000 current/torque limit  ->  SoE IDN S-0-0092 "Bipolar torque limit value".
    // *** MAP THESE AS PDO ***: add IDN 92 (hex #x005C, UINT16) to each drive's MDT,
    //   then link:  nMotor1_CurrentLimit_Raw -> Drive 1 (AX5112) S-0-0092
    //               nMotor2_CurrentLimit_Raw -> Drive 2 (AX5125) S-0-0092
    // Raw = 0.1 % per LSB (1000 = 100.0 %); scaled from stMotorX_Cmd.fCurrentLimit_pct
    // in PRG_Motion. Bipolar (limits both +/- torque), active in position mode (11).
    nMotor1_CurrentLimit_Raw AT %Q* : UINT;
    nMotor2_CurrentLimit_Raw AT %Q* : UINT;
END_VAR

// ---- GVLs/GVL_MenteeFoe.TcGVL
// Mentee V3.2 config-over-FoE command channel (FB_MenteeFoeFlash / PRG_Motion).
// The app writes the mtb_config_tool "config.bin" bytes into aData + nLen and
// pulses bExecute; the FB sends them to the motor slave over FoE (File access
// over EtherCAT), and — only on a validated download — writes CoE 0x1010:01
// = "save" so the firmware persists to flash and self-resets.
//
// config.bin = 32-byte header (magic 0x4D4F5452 / size / CRC32-IEEE) + payload
// (<= sizeof(Obj.params), max 2048). So the file is <= 2080 bytes. The app
// validates the header before writing here; the slave re-validates during FoE.
VAR_GLOBAL
    // ── command (written by the app over ADS) ──
    aData       : ARRAY[0..2079] OF BYTE;   // config.bin bytes (header + payload)
    nLen        : UDINT;                     // number of valid bytes in aData
    bExecute    : BOOL;                      // rising edge -> run FoE download (+ auto-save on success)

    // ── status (read by the app) ──
    nState      : INT;      // 0 IDLE | 1 OPEN | 2 WRITE | 3 CLOSE | 4 SAVE | 5 DONE | 6 ERROR
    bBusy       : BOOL;      // a flash sequence is in progress
    bDownloadOk : BOOL;      // FoE transfer accepted + validated by the slave (BEFORE the save)
    bDone       : BOOL;      // save command sent OK -> motor is self-resetting with the new config
    bError      : BOOL;      // sequence failed
    nErrId      : UDINT;     // ADS/FoE/CoE error id (when bError)
    nStage      : UDINT;     // stage that failed: 1 open | 2 write | 3 close | 4 save
END_VAR

// ---- GVLs/GVL_Encoder.TcGVL
{attribute 'TcGvlVarFlags' := 'OPC'}
VAR_GLOBAL
    // EL5112 encoder data — written by FB_EncoderHandler, read by Python over ADS
    // ADS symbol: GVL_Encoder.stEncoder
    stEncoder1          : ST_EncoderData;
    stEncoder2          : ST_EncoderData;

    // Encoder scaling — set once from Python or MAIN
    // fCountsPerUnit: how many encoder counts = 1 engineering unit
    // Example: 4096 counts/rev with units in degrees → fCountsPerUnit = 4096/360
    fCountsPerUnit1     : LREAL := 1.0;
    fCountsPerUnit2     : LREAL := 1.0;
END_VAR

// ---- GVLs/GVL_IO.TcGVL
{attribute 'qualified_only'}
VAR_GLOBAL
	RedLED 			  AT %Q*: BOOL;
	GreenLED 		  AT %Q*: BOOL;
	BlueLED			  AT %Q*: BOOL;
	b_MotorCooling			  AT %Q*: BOOL;
	    // I/O module state — Python can read inputs and write output setpoints
    // ADS symbol: GVL_IO.stIO
    stIO            : ST_IOData;

END_VAR

// ---- GVLs/GVL_MenteeMotor.TcGVL
{attribute 'TcGvlVarFlags' := 'OPC'}
VAR_GLOBAL
    // Commands — written by Python over ADS, sent to device every cycle
    // ADS symbol: GVL_MenteeMotor.stCmd
    stCmd               : ST_MenteeMotorCmd;

    // Status — read from device every cycle, read by Python over ADS
    // ADS symbol: GVL_MenteeMotor.stStatus
    stStatus            : ST_MenteeMotorStatus;
END_VAR

// ---- GVLs/GVL_MenteeMotorV32_OS.TcGVL
{attribute 'TcGvlVarFlags' := 'OPC'}
VAR_GLOBAL
    // ADS symbol: GVL_MenteeMotorV32_OS.stCmd
    stCmd    : ST_MenteeMotorV32OsCmd;
    // ADS symbol: GVL_MenteeMotorV32_OS.stStatus
    stStatus : ST_MenteeMotorV32OsStatus;

    // EtherCAT AL state of the Motor Slave V3.2 ("Box 1 (Motor Slave)").
    // >>> LINK IN XAE: <Motor Slave> > InfoData > State  ->  this variable. <<<
    // The EtherCAT master updates it every cycle (no ADS/FB needed). Decode:
    // low nibble = AL state (1=INIT, 2=PREOP, 4=SAFEOP, 8=OP), bit 4 = error.
    nSlaveState AT %I* : UINT;

    // V3.2 motion-profile command/status (FB_TrajectoryGen). The app writes the
    // params + pulses bStart; the FB streams the profile at 1 kHz into stCmd.
    // ADS symbol: GVL_MenteeMotorV32_OS.stTraj
    stTraj   : ST_MenteeTrajCmd;
END_VAR

// ---- GVLs/GVL_Profiles.TcGVL
{attribute 'TcGvlVarFlags' := 'OPC'}
// Synchronized motion-profile coordination. The app configures each enabled half
// (the Mentee profile lives in GVL_MenteeMotorV32_OS.stTraj; the load motors here)
// then pulses ONE bStartSync. PRG_Motion detects its rising edge and starts every
// enabled half in the SAME PLC cycle -> cycle-accurate (<=1 ms) synchronization,
// because all generators run in the same task at the same fTaskCycleS.
VAR_GLOBAL
    // Load-motor profiles (Beckhoff AX5000), one per axis.
    // ADS: GVL_Profiles.stLoadProfile1 / .stLoadProfile2
    stLoadProfile1 : ST_LoadProfileCmd;   // Motor 1 (Axis1)
    stLoadProfile2 : ST_LoadProfileCmd;   // Motor 2 (Axis2)

    // Mentee half participates in the synchronized start (its config + params are
    // in GVL_MenteeMotorV32_OS.stTraj; this only gates the shared start edge).
    // ADS: GVL_Profiles.bMenteeEnable
    bMenteeEnable  : BOOL;

    // Shared start/stop. Pulse bStartSync (rising edge) AFTER writing all enabled
    // halves' configs; PRG_Motion arms every enabled half that same cycle.
    // ADS: GVL_Profiles.bStartSync / .bStopSync
    bStartSync     : BOOL;
    bStopSync      : BOOL;
END_VAR

// ---- GVLs/GVL_CsvProfile.TcGVL
{attribute 'TcGvlVarFlags' := 'OPC'}
// Generic CSV-trajectory profile. The app uploads the resampled, unit-converted
// sample arrays + config into stCsv, then pulses stCsv.bStart; FB_CsvPlayer
// (called in PRG_Motion) replays it at the task rate, synchronized across both
// motors. Read/written GUARDED by the app (a PLC image without GVL_CsvProfile must
// not break the rest of telemetry).
VAR_GLOBAL
    // ADS: GVL_CsvProfile.stCsv (buffers written in chunks: stCsv.aMentee / .aLoad)
    stCsv : ST_CsvProfile;
END_VAR

// ---- GVLs/GVL_Slot2.TcGVL
{attribute 'TcGvlVarFlags' := 'OPC'}
// Generic slot-2 debug-PDO pipe coordination (new Mentee 3.2 pipeline).
// The app writes stCfg (binding addresses from the FW build's .map/.elf) and pulses
// bConfigure; FB_Slot2PipeHandler binds the lanes/slots and then runs the pipe,
// presenting the SAME ST_MenteeMotorV32OsCmd/Status contract as the legacy fixed pipe
// (GVL_MenteeMotorV32_OS) so profiles/CSV/recorder/GUI stay unchanged above it.
// FSM/main/mode commands go via CoE SDO 0x2000:01 (FB_MenteeSdoCmd) — the debug RxPDO
// has no control word.
VAR_GLOBAL
    // ── binding configuration (app -> PLC) ─────────────────────────────
    stCfg        : ST_Slot2Cfg;
    bConfigure   : BOOL;      // rising edge -> CLEAR_ALL + walk stCfg bindings
    bClearAll    : BOOL;      // rising edge -> CLEAR_ALL only (pipe goes idle)

    // ── pipe status (PLC -> app) ───────────────────────────────────────
    nBindState   : BYTE;      // 0 idle | 1 clearing | 2 binding | 3 RUN | 4 error
    bPipeActive  : BOOL;      // TRUE = bindings applied, adapter running
    bBindError   : BOOL;      // a bind command was rejected (fault=1) or timed out
    nFailedSlot  : BYTE;      // which walk step failed (16#FF = none)
    nCaptureCount: UDINT;     // raw 0x6001:0x0A capture counter (new FW semantics)
    nVarCount    : UDINT;     // slave-reported bound monitor lanes
    nLastOp      : UDINT;     // slave op echo (diagnostics)
    nFault       : UDINT;     // slave fault echo (diagnostics)

    // ── CoE SDO command channel (app -> PLC -> slave 0x2000:01) ────────
    nSdoOpcode   : BYTE;      // ec_command_id_e opcode to send
    bSdoExecute  : BOOL;      // rising edge -> send nSdoOpcode
    bSdoBusy     : BOOL;
    bSdoDone     : BOOL;      // last send completed OK (cleared on next execute)
    bSdoError    : BOOL;
    nSdoErrId    : UDINT;     // ADS error from FB_EcCoESdoWrite
END_VAR

// ---- GVLs/GVL_Recording.TcGVL
{attribute 'TcGvlVarFlags' := 'OPC'}
// High-rate recording: PLC fills a ring of chunks at the task rate; the app
// bulk-reads completed chunks over ADS and writes them to a file.
//
// HANDSHAKE (all ADS symbols under GVL_Recording.*):
//   app  -> bEnable    : start/stop recording (rising edge resets the ring)
//   app  -> nAckSeq    : last chunk sequence the app has fully read (overflow calc)
//   PLC  -> nChunkSeq  : completed-chunk counter (bumped each time a chunk fills)
//   PLC  -> nReadyIdx   : ring slot of the most recently completed chunk (0..REC_RING-1)
//   PLC  -> nDropped    : frames lost because the app fell behind (should stay 0)
//   PLC  -> aChunks     : the chunk ring (read aChunks[nReadyIdx].* per channel)
//
// The app reads a COMPLETED chunk (one the FB has already advanced past), so with
// REC_RING slots it has (REC_RING-1)*REC_CHUNK/rate seconds to read before the FB
// laps back to that slot — REC_RING-1 chunks of read slack (REC_CHUNK frames each).
VAR_GLOBAL CONSTANT
    REC_CHUNK      : UDINT := 2000;   // EtherCAT frames per chunk (chunk period = REC_CHUNK / task-rate)
    REC_RING       : UDINT := 4;      // number of chunks in the ring (read slack)
    REC_OVERSAMPLE : UDINT := 10;     // Mentee oversamples per frame — MUST match firmware OVERSAMPLE_SAMPLES_PER_CYCLE
    REC_FUTEK_OS   : UDINT := 5;      // Futek analog oversamples per frame (EL3702 x5) — MUST match ST_AnalogInData nChx_Sample len
END_VAR

VAR_GLOBAL
    // ── control (app writes) ──
    bEnable   : BOOL;     // TRUE = recording; rising edge clears the ring + counters
    nAckSeq   : UDINT;    // last chunk seq the app finished reading

    // ── status (PLC writes, app reads) ──
    nChunkSeq : UDINT;    // completed-chunk counter (monotonic; 0 = none yet this session)
    nReadyIdx : BYTE;     // ring slot of the most recently completed chunk
    nDropped  : UDINT;    // frames dropped (app too slow / overflow) — should remain 0
    bRunning  : BOOL;     // echoes bEnable once latched (diagnostic)

    // ── the chunk ring (ADS-read per channel array) ──
    aChunks   : ARRAY[0..REC_RING - 1] OF ST_RecChunk;
END_VAR

// ---- GVLs/GVL_Safety.TcGVL
{attribute 'qualified_only'}
VAR_GLOBAL
	//ST_TwinSAFE_IN
	stTwinSAFE_OUT	AT %Q* :ST_TwinSAFE_OUT;
	stTwinSAFE_IN	AT %I* : ST_TwinSAFE_IN;
	DoorMonitorFromPLC AT %I* : BOOL;
	SolonoidStatus AT %I* : BOOL;
END_VAR

// ---- GVLs/GVL_Status.TcGVL
{attribute 'TcGvlVarFlags' := 'OPC'}
VAR_GLOBAL
    // Status structs written by PLC every cycle, read by Python over ADS
    // ADS symbol: GVL_Status.stMotor1_Status
    //             GVL_Status.stMotor2_Status
    stMotor1_Status : ST_MotorStatus;
    stMotor2_Status : ST_MotorStatus;
END_VAR

// ---- GVLs/GVL_Sync.TcGVL
VAR_GLOBAL
    // Synchronized snapshot — all data from the same DC cycle.
    // Read from Python via single ADS read: GVL_Sync.stSnapshot
    stSnapshot : ST_SyncSnapshot;
END_VAR

// ---- GVLs/GVL_UartBridge.TcGVL
{attribute 'TcGvlVarFlags' := 'OPC'}
VAR_GLOBAL
    // Commands — written by Python over ADS, sent to device every cycle
    // ADS symbol: GVL_UartBridge.stCmd
    stCmd               : ST_UartBridgeCmd;

    // Status — read from device every cycle, read by Python over ADS
    // ADS symbol: GVL_UartBridge.stStatus
    stStatus            : ST_UartBridgeStatus;
END_VAR

// ---- POUs/MAIN.TcPOU
PROGRAM MAIN
VAR
	i: INT;
	ton_TwinSAFE_ACK_reset: TON;
	BlinkLED: ton;

	Pulse_On_TON: TON;
	Pulse_Off_TON: TON;
	bPulse	:	BOOL	;
	
	t_BlinkTime : TIME	;
	
	n_SafeSate	:	INT	;
END_VAR

i:=i+1;


ton_TwinSAFE_ACK_reset(IN:=GVL_Safety.stTwinSAFE_OUT.ErrACK, PT:=T#10S);
IF ton_TwinSAFE_ACK_reset.Q THEN;
	GVL_Safety.stTwinSAFE_OUT.ErrACK:=FALSE;
END_IF
GVL_Safety.stTwinSAFE_OUT.DoorMonitor:=GVL_Safety.DoorMonitorFromPLC;

//Battery Relay CMD
IF GVL_Safety.stTwinSAFE_OUT.BatRelay_CMD THEN
	GVL_Safety.stTwinSAFE_OUT.BatRelay_Manual_Off:=FALSE;
	GVL_Safety.stTwinSAFE_OUT.BatRelay_Manual_On:=TRUE;
ELSE
	GVL_Safety.stTwinSAFE_OUT.BatRelay_Manual_Off:=TRUE;
	GVL_Safety.stTwinSAFE_OUT.BatRelay_Manual_On:=FALSE;
END_IF

//Battery BMS Relay CMD
IF GVL_Safety.stTwinSAFE_OUT.BatBMS_Cmd THEN
	GVL_Safety.stTwinSAFE_OUT.RB_BatBMS_Manual_Off:=FALSE;
	GVL_Safety.stTwinSAFE_OUT.RB_BatBMS_Manual_On:=TRUE;
ELSE
	GVL_Safety.stTwinSAFE_OUT.RB_BatBMS_Manual_Off:=TRUE;
	GVL_Safety.stTwinSAFE_OUT.RB_BatBMS_Manual_On:=FALSE;

END_IF

act_LED_Control();
act_LogicMap();

ACTION act_LED_Control:
//Red 
IF GVL_Safety.stTwinSAFE_IN.EStop_Ok AND GVL_Safety.stTwinSAFE_IN.EStop_Status THEN
	//Red Off
	GVL_IO.RedLED:= FALSE;
ELSIF GVL_Safety.stTwinSAFE_IN.EStop_Ok=FALSE AND GVL_Safety.stTwinSAFE_IN.EStop_Status  THEN
	//Red Blink 
	GVL_IO.RedLED:=bPulse;
ELSIF GVL_Safety.stTwinSAFE_IN.EStop_Ok=FALSE AND GVL_Safety.stTwinSAFE_IN.EStop_Status=FALSE THEN
	//Red On
	GVL_IO.RedLED:= TRUE;
END_IF

//Blue
IF (GVL_Safety.stTwinSAFE_OUT.DoorMonitor AND GVL_Safety.stTwinSAFE_IN.Speps.step1) 
OR (GVL_Safety.stTwinSAFE_OUT.DoorMonitor=FALSE AND GVL_Safety.stTwinSAFE_IN.Speps.stepRnD) THEN
	//Blue Blink
	GVL_IO.BlueLED:=bPulse;
ELSIF GVL_Safety.stTwinSAFE_OUT.DoorMonitor AND GVL_Safety.stTwinSAFE_OUT.SolenoedMonitor=FALSE AND NOT GVL_Safety.stTwinSAFE_IN.Speps.stepRnD THEN
	//Blue Off
	GVL_IO.BlueLED:=FALSE;
ELSIF GVL_Safety.stTwinSAFE_OUT.DoorMonitor=FALSE OR (GVL_Safety.stTwinSAFE_IN.Speps.stepRnD AND GVL_Safety.stTwinSAFE_OUT.DoorMonitor) THEN
	//Blue On
	GVL_IO.BlueLED:=TRUE;
END_IF

//Green
IF (GVL_Safety.stTwinSAFE_IN.Speps.step1 AND GVL_Safety.stTwinSAFE_IN.EStop_Ok AND GVL_Safety.stTwinSAFE_OUT.DoorMonitor=TRUE) OR GVL_Safety.stTwinSAFE_IN.TransitionStep THEN
	//Green Blink
	GVL_IO.GreenLED:=bPulse;
ELSIF GVL_Safety.stTwinSAFE_IN.Safety_Armed OR (GVL_Safety.stTwinSAFE_IN.Speps.stepRnD) OR GVL_Safety.stTwinSAFE_IN.Speps.step2 THEN
	//Green On
	GVL_IO.GreenLED:=TRUE;
ELSIF GVL_Safety.stTwinSAFE_IN.Speps.step4 OR GVL_Safety.stTwinSAFE_IN.Speps.step5 
OR GVL_Safety.stTwinSAFE_IN.Speps.step6 OR GVL_Safety.stTwinSAFE_OUT.DoorMonitor=FALSE THEN
	//Green Off
	GVL_IO.GreenLED:=FALSE;
END_IF

IF GVL_Safety.stTwinSAFE_IN.Speps.step2 OR GVL_Safety.stTwinSAFE_IN.TransitionStep THEN
	t_BlinkTime:=T#0.5S;
ELSE
	t_BlinkTime:=T#1.5S;
END_IF

Pulse_On_TON(IN:=NOT bPulse , PT:=t_BlinkTime , Q=> , ET=> );
Pulse_Off_TON(IN:=bPulse , PT:=t_BlinkTime , Q=> , ET=> );
IF Pulse_On_TON.Q AND NOT bPulse THEN bPulse:=TRUE; END_IF;
IF Pulse_Off_TON.Q AND bPulse THEN bPulse:=FALSE; END_IF;


GVL_Safety.stTwinSAFE_IN.HV_Healthy_Invert:=NOT GVL_Safety.stTwinSAFE_IN.HV_Healthy;
GVL_Safety.stTwinSAFE_IN.LV_Healthy_Invert:=NOT GVL_Safety.stTwinSAFE_IN.LV_Healthy;
END_ACTION

ACTION act_LogicMap:
(*
_________________________________________________________________________________________________________________________________________________________________
Function				|	Bit 1 (RnD Mode) GVL_Safety.stTwinSAFE_OUT.Set_RnD_Mode		|	Bit 2 (RnD Mode 2)		GVL_Safety.stTwinSAFE_OUT.Set_RnD_Mode2	|
________________________|_______________________________|_______________________________|
From Safe to RnD		|	1							|	0							|
________________________|_______________________________|_______________________________|
From RnD to Armed		|	1							|	1							|
________________________|_______________________________|_______________________________|
From RnD to Safe		|	0							|	0							|
________________________|_______________________________|_______________________________|
From Armed to RnD		|	0							|	1							|
________________________|_______________________________|_______________________________|

*)
;

GVL_Safety.stTwinSAFE_OUT.Set_RnD_Mode;
GVL_Safety.stTwinSAFE_OUT.Set_RnD_Mode2;

CASE n_SafeSate OF
	E_SafetyState.enum_RnD_2_Safe://From RnD to Safe	
		GVL_Safety.stTwinSAFE_OUT.Set_RnD_Mode:=FALSE;
		GVL_Safety.stTwinSAFE_OUT.Set_RnD_Mode2:=FALSE;
	E_SafetyState.enum_Safe_2_RnD://From Safe to RnD
		GVL_Safety.stTwinSAFE_OUT.Set_RnD_Mode:=TRUE;
		GVL_Safety.stTwinSAFE_OUT.Set_RnD_Mode2:=FALSE;
	
	E_SafetyState.enum_RnD_2_Armed://From RnD to Armed
		GVL_Safety.stTwinSAFE_OUT.Set_RnD_Mode:=TRUE;
		GVL_Safety.stTwinSAFE_OUT.Set_RnD_Mode2:=TRUE;
	
	E_SafetyState.enum_Armed_2_RnD://From Armed to RnD
		GVL_Safety.stTwinSAFE_OUT.Set_RnD_Mode:=TRUE;
		GVL_Safety.stTwinSAFE_OUT.Set_RnD_Mode2:=FALSE;
END_CASE


(*IF GVL_Safety.stTwinSAFE_OUT.Bypass_C1C2 THEN
	
END_IF*)
END_ACTION

END_PROGRAM

// ---- POUs/PRG_Motion.TcPOU
PROGRAM PRG_Motion
VAR
    //--- Position/velocity control (one per motor) ---
    fbMotor1        : FB_MotorControl;
    fbMotor2        : FB_MotorControl;

    //--- Torque control (one per motor) ---
    fbTorque1       : FB_TorqueControl;
    fbTorque2       : FB_TorqueControl;

    //--- I/O handler ---
    fbIO            : FB_IOHandler;

    //--- Encoder handler ---
    fbEncoder1      : FB_EncoderHandler;
    fbEncoder2      : FB_EncoderHandler;

    //--- Analog input handler ---
    fbAnalogIn1     : FB_AnalogInHandler;
    fbAnalogIn2     : FB_AnalogInHandler;

    //--- Mentee Motor Slave handler (V3.2, slot-1 simple PDO 0x1600/0x1A00) ---
    fbMenteeMotor   : FB_MenteeMotorHandler;

    //--- Mentee Motor V3.2 slot-2: GENERIC DEBUG-PDO PIPE (new pipeline; replaces the
    //    legacy fixed oversample handler — same GVL contract, new transport). FSM/mode
    //    commands ride CoE SDO 0x2000 via fbMenteeSdo (GVL_Slot2 request channel). ---
    fbSlot2Pipe         : FB_Slot2PipeHandler;
    fbMenteeSdo         : FB_MenteeSdoCmd;
    //--- Mentee config-over-FoE flash (config.bin -> slave, then CoE save-to-flash) ---
    fbMenteeFoe         : FB_MenteeFoeFlash;

    //--- Mentee Motor V3.2 trajectory generator (1 kHz trapezoid) ---
    fbMenteeTraj        : FB_TrajectoryGen;

    //--- Load-motor (Beckhoff) profile generators, synchronized with the Mentee
    //    profile via GVL_Profiles.bStartSync (torque waveform or ext-setpoint pos/vel) ---
    fbLoadProfile1      : FB_LoadMotorProfile;
    fbLoadProfile2      : FB_LoadMotorProfile;

    //--- Generic CSV-trajectory player (uploaded buffer; both motors synchronized) ---
    fbCsvPlayer         : FB_CsvPlayer;

    //--- High-rate recorder (buffers every frame into GVL_Recording.aChunks) ---
    fbRecorder          : FB_HighRateRecorder;

    //--- Mentee UART Bridge handler (V3.1) ---
    fbUartBridge    : FB_UartBridgeHandler;

    //--- NC Axis references — link to NC axes in XAE ---
    Axis1           : AXIS_REF;
    Axis2           : AXIS_REF;

    //--- Safety ---
    bEStopActive    : BOOL;

    //--- Task cycle period [s], read live from the running task config so the
    //    trajectory generator timestep auto-tracks any PlcTask CycleTime change
    //    (1 ms <-> 250 us) with no code edit here. ---
    fTaskCycleS     : REAL;
END_VAR

//----------------------------------------------------------------------
// 1. SAFETY — runs before everything else
//----------------------------------------------------------------------
bEStopActive := GVL_IO.stIO.bDI_EmergencyStop;

IF bEStopActive THEN
    GVL_Commands.stMotor1_Cmd.bEnable := FALSE;
    GVL_Commands.stMotor2_Cmd.bEnable := FALSE;
    GVL_Commands.stMotor1_Cmd.bStop   := TRUE;
    GVL_Commands.stMotor2_Cmd.bStop   := TRUE;
END_IF

//----------------------------------------------------------------------
// 2. I/O HANDLER — fresh sensor data before motion FBs
//----------------------------------------------------------------------
fbIO(
    nRawDigitalIn    := GVL_IO.stIO.nDigitalInputs,
    nRawAnalogIn_Ch1 := GVL_IO.stIO.nAnalogIn_Raw_Ch1,
    nRawAnalogIn_Ch2 := GVL_IO.stIO.nAnalogIn_Raw_Ch2,
    stIO             := GVL_IO.stIO
);

//----------------------------------------------------------------------
// 3. ENCODER HANDLER
//----------------------------------------------------------------------
fbEncoder1(stEncoder := GVL_Encoder.stEncoder1, fCountsPerUnit := GVL_Encoder.fCountsPerUnit1);
fbEncoder2(stEncoder := GVL_Encoder.stEncoder2, fCountsPerUnit := GVL_Encoder.fCountsPerUnit2);

//----------------------------------------------------------------------
// 4. ANALOG INPUT HANDLER
//----------------------------------------------------------------------
fbAnalogIn1(stAnalogIn := GVL_AnalogIn.stAnalogIn1);
fbAnalogIn2(stAnalogIn := GVL_AnalogIn.stAnalogIn2);

//----------------------------------------------------------------------
// 5. MENTEE MOTOR SLAVE — V3.2, slot-1 (simple PDO 0x1600/0x1A00)
//----------------------------------------------------------------------
fbMenteeMotor(
    stCmd    := GVL_MenteeMotor.stCmd,
    stStatus := GVL_MenteeMotor.stStatus
);

//----------------------------------------------------------------------
// 5a. MENTEE V3.2 motion-profile generator (1 kHz: sine/trapezoid/step/
//     s-curve/ramp). While a profile runs it overrides the selected setpoint
//     field (by nField) BEFORE the handler below forwards stCmd to the RxPDO.
//     Measured position = latest OS sub-sample (anchor for position profiles).
//----------------------------------------------------------------------
// Live task cycle [s] from the running task config (100 ns units -> s), so the
// profile timestep auto-tracks PlcTask CycleTime (1 ms <-> 250 us) — no edit here.
fTaskCycleS := LREAL_TO_REAL(UDINT_TO_LREAL(_TaskInfo[GETCURTASKINDEXEX()].CycleTime) * 1.0E-7);
IF fTaskCycleS <= 0.0 THEN
    fTaskCycleS := 0.001;    // safety fallback if the system var reads 0
END_IF

fbMenteeTraj(
    stTraj       := GVL_MenteeMotorV32_OS.stTraj,
    fMeasuredPos := GVL_MenteeMotorV32_OS.stStatus.fLatestPos,  // decoded theta (REAL)
    fDt          := fTaskCycleS,   // auto-tracks the PlcTask cycle (1 ms / 250 us)
    bStartSync   := GVL_Profiles.bStartSync AND GVL_Profiles.bMenteeEnable,
    bStopSync    := GVL_Profiles.bStopSync
);
IF fbMenteeTraj.bRunning THEN
    // route by the FB's LATCHED field (nFieldOut) — the live stTraj.nField can
    // already hold the NEXT run's field while the app rewrites the config over
    // ADS, and routing by it would inject this run's value into the wrong lane
    CASE fbMenteeTraj.nFieldOut OF
        1:  GVL_MenteeMotorV32_OS.stCmd.impedance_p_des   := fbMenteeTraj.fSetpoint;
        2:  GVL_MenteeMotorV32_OS.stCmd.setpoint_velocity := fbMenteeTraj.fSetpoint;
        3:  GVL_MenteeMotorV32_OS.stCmd.setpoint_current  := fbMenteeTraj.fSetpoint;
    ELSE
        GVL_MenteeMotorV32_OS.stCmd.setpoint_position := fbMenteeTraj.fSetpoint;
    END_CASE
END_IF

//----------------------------------------------------------------------
// 5a2. CSV TRAJECTORY PLAYER (generic uploaded buffer, both motors synchronized).
//      Called here so its Mentee output reaches the RxPDO forward (5b) THIS cycle
//      and its Beckhoff torque override precedes torque control (9). For a Beckhoff
//      POS/VEL run the FB feeds the NC axis via external setpoint — the motor must
//      already be ENABLED/READY (its MC_Power is maintained from prior cycles by
//      fbMotor1/2 in 7/8). Mutually exclusive with the closed-form profiles.
//----------------------------------------------------------------------
fbCsvPlayer(
    stCsv     := GVL_CsvProfile.stCsv,
    AxisLoad1 := Axis1,
    AxisLoad2 := Axis2,
    fLoad1Pos := Axis1.NcToPlc.ActPos,
    fLoad2Pos := Axis2.NcToPlc.ActPos,
    fDt       := fTaskCycleS
);
// The CSV player and the closed-form generators are mutually exclusive by design;
// the guards below enforce it (the CSV player YIELDS) so that if a closed-form
// profile is somehow still running it keeps ownership of the shared command field
// instead of both writing it (last-write-wins glitch).
IF fbCsvPlayer.bRunning AND GVL_CsvProfile.stCsv.bMenteeEnable AND NOT fbMenteeTraj.bRunning THEN
    CASE GVL_CsvProfile.stCsv.nMenteeField OF
        1:  GVL_MenteeMotorV32_OS.stCmd.impedance_p_des   := fbCsvPlayer.fMenteeOut;
        2:  GVL_MenteeMotorV32_OS.stCmd.setpoint_velocity := fbCsvPlayer.fMenteeOut;
        3:  GVL_MenteeMotorV32_OS.stCmd.setpoint_current  := fbCsvPlayer.fMenteeOut;
    ELSE
        GVL_MenteeMotorV32_OS.stCmd.setpoint_position := fbCsvPlayer.fMenteeOut;
    END_CASE
END_IF
IF fbCsvPlayer.bRunning AND GVL_CsvProfile.stCsv.bLoadEnable
   AND (GVL_CsvProfile.stCsv.nLoadDomain = 0) THEN   // TORQUE domain -> override fTargetTorque
    IF (GVL_CsvProfile.stCsv.nLoadMotor = 1) AND NOT fbLoadProfile1.bRunning THEN
        GVL_Commands.stMotor1_Cmd.fTargetTorque := fbCsvPlayer.fLoadOut;
    ELSIF (GVL_CsvProfile.stCsv.nLoadMotor = 2) AND NOT fbLoadProfile2.bRunning THEN
        GVL_Commands.stMotor2_Cmd.fTargetTorque := fbCsvPlayer.fLoadOut;
    END_IF
END_IF

//----------------------------------------------------------------------
// 5b. MENTEE MOTOR V3.2 — slot-2 GENERIC DEBUG PIPE (new pipeline).
//     Same GVL contract as the legacy handler: stCmd setpoints stream via the
//     bound inject slots; stStatus (incl. synthesized status word + oversample
//     view) is rebuilt from the debug TxPDO. FSM/main/mode commands go via
//     fbMenteeSdo (CoE SDO 0x2000; GVL_Slot2 channel) — stCmd.nControlWord is
//     no longer consumed. Bindings: app writes GVL_Slot2.stCfg + bConfigure.
//----------------------------------------------------------------------
fbSlot2Pipe(
    stCmd    := GVL_MenteeMotorV32_OS.stCmd,
    stStatus := GVL_MenteeMotorV32_OS.stStatus
);
fbMenteeSdo();
fbMenteeFoe();   // FoE config.bin download + auto-save on success (GVL_MenteeFoe channel)

//----------------------------------------------------------------------
// 6. MENTEE UART BRIDGE — V3.1
//----------------------------------------------------------------------
fbUartBridge(
    stCmd    := GVL_UartBridge.stCmd,
    stStatus := GVL_UartBridge.stStatus
);

//----------------------------------------------------------------------
// 6. LIMIT SWITCH INTERLOCKS
//----------------------------------------------------------------------
IF GVL_IO.stIO.bDI_LimitPos_M1 AND GVL_Commands.stMotor1_Cmd.fTargetVelocity > 0 THEN
    GVL_Commands.stMotor1_Cmd.bStop := TRUE;
END_IF
IF GVL_IO.stIO.bDI_LimitNeg_M1 AND GVL_Commands.stMotor1_Cmd.fTargetVelocity < 0 THEN
    GVL_Commands.stMotor1_Cmd.bStop := TRUE;
END_IF
IF GVL_IO.stIO.bDI_LimitPos_M2 AND GVL_Commands.stMotor2_Cmd.fTargetVelocity > 0 THEN
    GVL_Commands.stMotor2_Cmd.bStop := TRUE;
END_IF
IF GVL_IO.stIO.bDI_LimitNeg_M2 AND GVL_Commands.stMotor2_Cmd.fTargetVelocity < 0 THEN
    GVL_Commands.stMotor2_Cmd.bStop := TRUE;
END_IF

//----------------------------------------------------------------------
// 7. MOTOR 1
//----------------------------------------------------------------------
fbMotor1(
    Axis     := Axis1,
    stCmd    := GVL_Commands.stMotor1_Cmd,
    stStatus => GVL_Status.stMotor1_Status
);

GVL_IO.stIO.bDO_BrakeRelease_M1 :=
    (GVL_Status.stMotor1_Status.eState = E_MotorState.READY)  OR
    (GVL_Status.stMotor1_Status.eState = E_MotorState.MOVING) OR
    (GVL_Status.stMotor1_Status.eState = E_MotorState.HOMING);

//----------------------------------------------------------------------
// 8. MOTOR 2
//----------------------------------------------------------------------
fbMotor2(
    Axis     := Axis2,
    stCmd    := GVL_Commands.stMotor2_Cmd,
    stStatus => GVL_Status.stMotor2_Status
);

GVL_IO.stIO.bDO_BrakeRelease_M2 :=
    (GVL_Status.stMotor2_Status.eState = E_MotorState.READY)  OR
    (GVL_Status.stMotor2_Status.eState = E_MotorState.MOVING) OR
    (GVL_Status.stMotor2_Status.eState = E_MotorState.HOMING);
	
//----------------------------------------------------------------------
// 8b. CURRENT / TORQUE LIMIT  ->  AX5000 SoE S-0-0092 (mapped MDT PDO)
//     % setpoint -> raw IDN units. 0.1 % per LSB => 1000 = 100.0 %.
//     VERIFY the S-0-0092 weighting in Drive Manager; if it is 0.01 %, use 100.0.
//     NOTE: 0 % = no torque -> the axis cannot hold or move.
//----------------------------------------------------------------------
GVL_Commands.nMotor1_CurrentLimit_Raw :=
    LREAL_TO_UINT(LIMIT(0.0, GVL_Commands.stMotor1_Cmd.fCurrentLimit_pct, 100.0) * 10.0);
GVL_Commands.nMotor2_CurrentLimit_Raw :=
    LREAL_TO_UINT(LIMIT(0.0, GVL_Commands.stMotor2_Cmd.fCurrentLimit_pct, 100.0) * 10.0);

//----------------------------------------------------------------------
// 8c. LOAD-MOTOR PROFILES (Beckhoff) — synchronized with the Mentee profile via
//     GVL_Profiles.bStartSync. Placed AFTER MC_Power (so the external-setpoint
//     feed acts on an already-powered axis) and BEFORE torque control (so a
//     TORQUE-domain profile overrides fTargetTorque before FB_TorqueControl
//     streams it). fMeasuredPos = axis actual position [deg] for anchoring.
//       nDomain 0 TORQUE  : override stMotorN_Cmd.fTargetTorque while running.
//                           The app must already be in torque mode
//                           (eControlMode=TORQUE, bTorqueExecute=TRUE).
//       nDomain 1/2 POS/VEL: the FB feeds the NC axis via external setpoint; the
//                           motor must be ENABLED/READY and NOT executing a move.
//----------------------------------------------------------------------
fbLoadProfile1(
    stProfile    := GVL_Profiles.stLoadProfile1,
    Axis         := Axis1,
    fMeasuredPos := Axis1.NcToPlc.ActPos,
    fDt          := fTaskCycleS,
    bStartSync   := GVL_Profiles.bStartSync,
    bStopSync    := GVL_Profiles.bStopSync
);
IF fbLoadProfile1.bRunning AND (GVL_Profiles.stLoadProfile1.nDomain = 0) THEN
    GVL_Commands.stMotor1_Cmd.fTargetTorque := fbLoadProfile1.fSetpoint;
END_IF

fbLoadProfile2(
    stProfile    := GVL_Profiles.stLoadProfile2,
    Axis         := Axis2,
    fMeasuredPos := Axis2.NcToPlc.ActPos,
    fDt          := fTaskCycleS,
    bStartSync   := GVL_Profiles.bStartSync,
    bStopSync    := GVL_Profiles.bStopSync
);
IF fbLoadProfile2.bRunning AND (GVL_Profiles.stLoadProfile2.nDomain = 0) THEN
    GVL_Commands.stMotor2_Cmd.fTargetTorque := fbLoadProfile2.fSetpoint;
END_IF

//----------------------------------------------------------------------
// 9. TORQUE CONTROL
//----------------------------------------------------------------------
fbTorque1(Axis := Axis1, stCmd := GVL_Commands.stMotor1_Cmd,
          bAxisReady := (GVL_Status.stMotor1_Status.eState = E_MotorState.READY));
GVL_Status.stMotor1_Status.bTorqueActive   := fbTorque1.stStatus.bTorqueActive;
GVL_Status.stMotor1_Status.bTorqueInTorque := fbTorque1.stStatus.bTorqueInTorque;
IF fbTorque1.stStatus.bError THEN
    GVL_Status.stMotor1_Status.bError   := TRUE;
    GVL_Status.stMotor1_Status.nErrorID := fbTorque1.stStatus.nErrorID;
END_IF

fbTorque2(Axis := Axis2, stCmd := GVL_Commands.stMotor2_Cmd,
          bAxisReady := (GVL_Status.stMotor2_Status.eState = E_MotorState.READY));
GVL_Status.stMotor2_Status.bTorqueActive   := fbTorque2.stStatus.bTorqueActive;
GVL_Status.stMotor2_Status.bTorqueInTorque := fbTorque2.stStatus.bTorqueInTorque;
IF fbTorque2.stStatus.bError THEN
    GVL_Status.stMotor2_Status.bError   := TRUE;
    GVL_Status.stMotor2_Status.nErrorID := fbTorque2.stStatus.nErrorID;
END_IF

//----------------------------------------------------------------------
// 10. STATUS LEDs
//----------------------------------------------------------------------
GVL_IO.stIO.bDO_StatusLED_Green :=
    NOT GVL_Status.stMotor1_Status.bError AND
    NOT GVL_Status.stMotor2_Status.bError AND
    NOT bEStopActive;

GVL_IO.stIO.bDO_StatusLED_Red :=
    GVL_Status.stMotor1_Status.bError OR
    GVL_Status.stMotor2_Status.bError OR
    bEStopActive;

//----------------------------------------------------------------------
// 11. SYNCHRONIZED SNAPSHOT — all data from this DC cycle
//     Python reads GVL_Sync.stSnapshot in a single ADS call.
//     nCycleCount lets Python detect missed or duplicate reads.
//----------------------------------------------------------------------
GVL_Sync.stSnapshot.nCycleCount     := GVL_Sync.stSnapshot.nCycleCount + 1;
GVL_Sync.stSnapshot.nDcTimestamp    := F_GetCurDcTaskTime64();

// UART Bridge (V3.1)
GVL_Sync.stSnapshot.stBridge        := GVL_UartBridge.stStatus;

// Mentee Motor (V3.2, slot-1)
GVL_Sync.stSnapshot.stMotor         := GVL_MenteeMotor.stStatus;

// Mentee Motor (V3.2, slot-2 oversample)
GVL_Sync.stSnapshot.stMotorV32_OS   := GVL_MenteeMotorV32_OS.stStatus;
// EtherCAT AL state (Motor Slave InfoData.State, linked to nSlaveState) — the
// master's authoritative online view: (nAlState AND 16#000F) = 8 means OP.
GVL_Sync.stSnapshot.stMotorV32_OS.nAlState := GVL_MenteeMotorV32_OS.nSlaveState;
// V3.2 trajectory generator running flag (so the app can reflect it).
GVL_Sync.stSnapshot.bTrajRunning := fbMenteeTraj.bRunning;

// Encoders
GVL_Sync.stSnapshot.stEncoder1      := GVL_Encoder.stEncoder1;
GVL_Sync.stSnapshot.stEncoder2      := GVL_Encoder.stEncoder2;

// Analog inputs
GVL_Sync.stSnapshot.stAnalogIn1     := GVL_AnalogIn.stAnalogIn1;
GVL_Sync.stSnapshot.stAnalogIn2     := GVL_AnalogIn.stAnalogIn2;

// Motor control status
GVL_Sync.stSnapshot.stMotor1Status  := GVL_Status.stMotor1_Status;
GVL_Sync.stSnapshot.stMotor2Status  := GVL_Status.stMotor2_Status;

// Safety
GVL_Sync.stSnapshot.bEStopActive    := bEStopActive;

//----------------------------------------------------------------------
// 12. HIGH-RATE RECORDER — append this frame to the recording ring while
//     GVL_Recording.bEnable. Runs last, on the freshly-assembled snapshot.
//----------------------------------------------------------------------
fbRecorder(stSnap := GVL_Sync.stSnapshot);

END_PROGRAM

// ---- POUs/FB_MotorControl.TcPOU
FUNCTION_BLOCK FB_MotorControl
VAR_IN_OUT
    Axis            : AXIS_REF;
END_VAR

VAR_INPUT
    stCmd           : ST_MotorCommand;
END_VAR

VAR_OUTPUT
    stStatus        : ST_MotorStatus;
END_VAR

VAR
    nActTorque_Raw  AT %I* : INT;

    fbPower         : MC_Power;
    fbMoveAbs       : MC_MoveAbsolute;
    fbMoveRel       : MC_MoveRelative;
    fbMoveVel       : MC_MoveVelocity;
    fbStop          : MC_Stop;
    fbReset         : MC_Reset;
    fbSoeReset      : FB_SoEReset;     // Tc2_MC2_Drive — SoE drive reset (S-0-0099)
    fbHome          : MC_Home;
    fbSetPosition   : MC_SetPosition;

    rtExecuteMove   : R_TRIG;
    rtStop          : R_TRIG;
    rtResetError    : R_TRIG;
    rtSoeReset      : R_TRIG;          // diagnostic: SoE drive reset only
    rtNcReset       : R_TRIG;          // diagnostic: NC axis reset only
    rtHome          : R_TRIG;
    rtZeroPosition  : R_TRIG;
    ftSoeBusy       : F_TRIG;          // SoE-reset Busy falling edge -> clear the latch

    eState          : E_MotorState;
    bMoveLatch      : BOOL;
    bSoeResetExec   : BOOL;            // latch: SoE drive reset requested / in progress
    bNcResetExec    : BOOL;            // latch: NC axis reset requested / in progress
    nResetStage     : BYTE;            // RESETTING sequence: 1 SoE | 2 settle | 3 NC
    tonSettle       : TON;             // drive-settle gap between SoE and NC reset
    tonResetGuard   : TON;             // whole-sequence watchdog -> back to ERROR
    fPrevVelocity   : LREAL;
END_VAR
VAR CONSTANT
    T_RESET_SETTLE  : TIME := T#250MS; // drive settle after the SoE reset completes
    T_RESET_GUARD   : TIME := T#15S;   // > FB_SoEReset's 10 s timeout + NC reset
END_VAR

//----------------------------------------------------------------------
// EDGE DETECTION
//----------------------------------------------------------------------
rtExecuteMove (CLK := stCmd.bExecuteMove);
rtStop        (CLK := stCmd.bStop);
rtResetError  (CLK := stCmd.bResetError);
rtSoeReset    (CLK := stCmd.bSoeReset);
rtNcReset     (CLK := stCmd.bNcReset);
rtHome        (CLK := stCmd.bHome);
rtZeroPosition(CLK := stCmd.bZeroPosition);

// Diagnostic single-shot resets — latch the respective background FB. Gated
// to non-motion states: MC_Reset on a MOVING axis hard-aborts the travel
// command (no deceleration ramp) and an SoE reset is comparably disruptive
// at the drive level — on a coupled bench that is a mechanical hazard, not a
// diagnostic. (The full sequenced recovery is the bResetError path below.)
IF (eState = E_MotorState.DISABLED) OR (eState = E_MotorState.READY)
        OR (eState = E_MotorState.ERROR) THEN
    IF rtSoeReset.Q THEN
        bSoeResetExec := TRUE;
    END_IF
    IF rtNcReset.Q THEN
        bNcResetExec := TRUE;
    END_IF
END_IF

//----------------------------------------------------------------------
// POWER — called every cycle
//----------------------------------------------------------------------
fbPower(
    Axis            := Axis,
    Enable          := (eState = E_MotorState.ENABLING
                     OR eState = E_MotorState.READY
                     OR eState = E_MotorState.MOVING
                     OR eState = E_MotorState.STOPPING
                     OR eState = E_MotorState.HOMING),
    Enable_Positive := (eState = E_MotorState.ENABLING
                     OR eState = E_MotorState.READY
                     OR eState = E_MotorState.MOVING
                     OR eState = E_MotorState.STOPPING
                     OR eState = E_MotorState.HOMING),
    Enable_Negative := (eState = E_MotorState.ENABLING
                     OR eState = E_MotorState.READY
                     OR eState = E_MotorState.MOVING
                     OR eState = E_MotorState.STOPPING
                     OR eState = E_MotorState.HOMING),
    Override        := 100.0,
    BufferMode      := MC_Aborting);

//----------------------------------------------------------------------
// SET POSITION — zero axis on rising edge, only in READY state
//----------------------------------------------------------------------
fbSetPosition(
    Axis     := Axis,
    Execute  := rtZeroPosition.Q,
    Position := 0.0,
    Mode     := FALSE);

IF fbSetPosition.Done  THEN stStatus.bZeroDone := TRUE; END_IF
IF fbSetPosition.Error THEN stStatus.bError    := TRUE;
                             stStatus.nErrorID  := fbSetPosition.ErrorID; END_IF

//----------------------------------------------------------------------
// STOP FB — called every cycle, Execute held TRUE only in STOPPING
//----------------------------------------------------------------------
fbStop(
    Axis         := Axis,
    Execute      := (eState = E_MotorState.STOPPING),
    Deceleration := SEL(stCmd.fDeceleration > 0, 500.0, stCmd.fDeceleration),
    Jerk         := stCmd.fJerk);

//----------------------------------------------------------------------
// MOVE FBs — called every cycle, Execute driven by state + latch
//----------------------------------------------------------------------
fbMoveAbs(
    Axis         := Axis,
    Execute      := bMoveLatch AND (eState = E_MotorState.MOVING)
                   AND (stCmd.eControlMode = E_ControlMode.POSITION)
                   AND NOT stCmd.bRelative,
    Position     := stCmd.fTargetPosition,
    Velocity     := SEL(stCmd.fTargetVelocity > 0,
                        stCmd.fMaxVelocity, stCmd.fTargetVelocity),
    Acceleration := stCmd.fAcceleration,
    Deceleration := stCmd.fDeceleration,
    Jerk         := stCmd.fJerk,
    BufferMode   := MC_Aborting);

fbMoveRel(
    Axis         := Axis,
    Execute      := bMoveLatch AND (eState = E_MotorState.MOVING)
                   AND (stCmd.eControlMode = E_ControlMode.POSITION)
                   AND stCmd.bRelative,
    Distance     := stCmd.fTargetPosition * stCmd.fDirection,
    Velocity     := SEL(stCmd.fTargetVelocity > 0,
                        stCmd.fMaxVelocity, stCmd.fTargetVelocity),
    Acceleration := stCmd.fAcceleration,
    Deceleration := stCmd.fDeceleration,
    Jerk         := stCmd.fJerk,
    BufferMode   := MC_Aborting);

fbMoveVel(
    Axis         := Axis,
    Execute      := bMoveLatch AND (eState = E_MotorState.MOVING)
                   AND (stCmd.eControlMode = E_ControlMode.VELOCITY),
    Velocity     := ABS(stCmd.fTargetVelocity),
    Direction    := SEL(stCmd.fTargetVelocity >= 0,
                        MC_Negative_Direction, MC_Positive_Direction),
    Acceleration := stCmd.fAcceleration,
    Deceleration := stCmd.fDeceleration,
    Jerk         := stCmd.fJerk,
    BufferMode   := MC_Aborting);

//----------------------------------------------------------------------
// SoE DRIVE RESET (FB_SoEReset, Tc2_MC2_Drive) — resets the AX5000 drive via
// S-0-0099 (a separate action from MC_Reset's NC reset). Called every cycle;
// triggered (latched) from the ERROR-state reset and runs to completion in the
// background. NetId '' = local controller; set it if the drive's NC is remote.
//----------------------------------------------------------------------
fbSoeReset(Axis := Axis, NetId := '', Execute := bSoeResetExec, Timeout := T#10S);
ftSoeBusy(CLK := fbSoeReset.Busy);
IF ftSoeBusy.Q THEN
    bSoeResetExec := FALSE;          // Busy 1->0: SoE reset finished (Error/SercosErrId valid)
END_IF
IF bSoeResetExec AND fbSoeReset.Error THEN
    bSoeResetExec := FALSE;          // immediate error (Busy never rose) -> don't hang the latch
END_IF

//----------------------------------------------------------------------
// NC AXIS RESET (MC_Reset) — called every cycle; latched from the sequenced
// recovery (RESETTING stage 3) or the diagnostic bNcReset command. The latch
// drops Execute back to FALSE on Done/Error, so every request produces a
// fresh rising edge (a one-shot Execute:=TRUE call would fire only once per
// PLC run — MC blocks trigger on the Execute edge).
//----------------------------------------------------------------------
fbReset(Axis := Axis, Execute := bNcResetExec);
IF bNcResetExec AND (fbReset.Done OR fbReset.Error) THEN
    bNcResetExec := FALSE;
END_IF

//----------------------------------------------------------------------
// STATE MACHINE
//----------------------------------------------------------------------
CASE eState OF

    E_MotorState.DISABLED:
        IF stCmd.bEnable THEN
            eState := E_MotorState.ENABLING;
        END_IF

    E_MotorState.ENABLING:
        IF NOT stCmd.bEnable THEN
            eState := E_MotorState.DISABLED;
        ELSIF fbPower.Error THEN
            eState := E_MotorState.ERROR;
        ELSIF fbPower.Status THEN
            eState := E_MotorState.READY;
        END_IF

    E_MotorState.READY:
        bMoveLatch    := FALSE;
        fPrevVelocity := 0.0;
        stCmd.bStop   := FALSE;

